// TIA Portal project "Projet Festo V4" (V20)

(* hardware
DEVICE "Station ET 200SP_1"  ET 200SP-Station
   slot 0: "Châssis_0"  Rack  6ES5 710-8MAx1
   slot 1: "6ES7512-1SK01-0AB0"  CPU 1512SP F-1 PN  6ES7 512-1SK01-0AB0  V2.8
      slot 32768: "Interface PROFINET_1"  X1
         slot 32771: "Port_3"  X1 P3
   slot 2: "F-DI 8x24VDC HF_1"  F-DI 8x24VDC HF  6ES7 136-6BA00-0CA0  V1.0
      slot 1: "F-DI 8x24VDC HF_1"  F-DI 8x24VDC HF
   slot 3: "F-DQ 4x24VDC/2A PM HF_1"  F-DQ 4x24VDC/2A PM HF  6ES7 136-6DB00-0CA0  V2.0
      slot 1: "F-DQ 4x24VDC/2A PM HF_1"  F-DQ 4x24VDC/2A PM HF
   slot 4: "F-RQ 1x24..48VDC/24..230VAC/5A_1"  F-RQ 1x24..48V DC/24..230VAC/5A  6ES7 136-6RA00-0BF0  V1.0
      slot 1: "F-RQ 1x24..48VDC/24..230VAC/5A_1"  F-RQ 1x24..48V DC/24..230VAC/5A
   slot 5: "DI 8x24VDC HF_1"  DI 8x24VDC HF  6ES7 131-6BF00-0CA0  V2.0
      slot 1: "DI 8x24VDC HF_1"  DI 8x24VDC HF
   slot 6: "DI 8x24VDC HF_2"  DI 8x24VDC HF  6ES7 131-6BF00-0CA0  V2.0
      slot 1: "DI 8x24VDC HF_2"  DI 8x24VDC HF
   slot 7: "DQ 8x24VDC/0.5A HF_1"  DQ 8x24VDC/0.5A HF  6ES7 132-6BF00-0CA0  V2.0
      slot 1: "DQ 8x24VDC/0.5A HF_1"  DQ 8x24VDC/0.5A HF
   slot 8: "DQ 8x24VDC/0.5A HF_2"  DQ 8x24VDC/0.5A HF  6ES7 132-6BF00-0CA0  V2.0
      slot 1: "DQ 8x24VDC/0.5A HF_2"  DQ 8x24VDC/0.5A HF
   slot 9: "AI 4xU/I 2-wire ST_1"  AI 4xU/I 2-wire ST  6ES7 134-6HD01-0BA1  V2.0
      slot 1: "AI 4xU/I 2-wire ST_1"  AI 4xU/I 2-wire ST
   slot 10: "AQ 4xU/I ST_1"  AQ 4xU/I ST  6ES7 135-6HD00-0BA1  V1.1
      slot 1: "AQ 4xU/I ST_1"  AQ 4xU/I ST
   slot 11: "Module serveur_1"  Server module  6ES7 193-6PA00-0AA0  V1.1
      slot 1: "Module serveur_1"  Server module
   slot 127: "BA 2xRJ45"  BA 2xRJ45  6ES7 193-6AR00-0AA0  V0.0
      slot 32769: "Port_1"  X1 P1  6ES7 193-6AR00-0AA0
      slot 32770: "Port_2"  X1 P2  6ES7 193-6AR00-0AA0
DEVICE "HMI_1"  MTP1000 Unified Comfort
   slot 0: "HMI_1"  MTP1000 Unified Comfort  6AV2 128-3KB06-0AXx  20.0.0.2
   slot 1: "HMI_RT_1"  MTP1000 Unified Comfort  6AV2 128-3KB06-0AXx  20.0.0.2
   slot 5: "HMI_1.IE_CP_1"  PROFINET Interface  20.0.0.2
      slot 1: "Interface PROFINET_1"  PROFINET Interface
         slot 1: "Port_1"  Port
         slot 2: "Port_2"  Port
   slot 6: "HMI_1.IE_CP_2"  PROFINET Interface  20.0.0.2
      slot 1: "Interface PROFINET_GBit"  PROFINET Interface
         slot 1: "Port_1"  Port
*)

// ===== PLC "6ES7512-1SK01-0AB0"  CPU 1512SP F-1 PN =====

VAR_GLOBAL   // PLC tag table "Table de variables standard"
   "Clock_Byte" AT %MB0 : Byte;   // Octet cadence B0
   "Clock_10Hz" AT %M0.0 : Bool;   // Octet cadence B0
   "Clock_5Hz" AT %M0.1 : Bool;   // Octet cadence B0
   "Clock_2.5Hz" AT %M0.2 : Bool;   // Octet cadence B0
   "Clock_2Hz" AT %M0.3 : Bool;   // Octet cadence B0
   "Clock_1.25Hz" AT %M0.4 : Bool;   // Octet cadence B0
   "Clock_1Hz" AT %M0.5 : Bool;   // Octet cadence B0
   "Clock_0.625Hz" AT %M0.6 : Bool;   // Octet cadence B0
   "Clock_0.5Hz" AT %M0.7 : Bool;   // Octet cadence B0
   "AURG_voie1" AT %I0.0 : Bool;   // Entrée Safety AURG
   "AURG_voie2" AT %I0.4 : Bool;   // Entrée Safety AURG
   "bouton_bleu" AT %I0.1 : Bool;   // acquittement apres AURG
   "voyant_bleu" AT %Q6.0 : Bool;   // Sortie Safety
   "FQ1" AT %Q6.1 : Bool;   // Sortie Safety pour relais
   "FQ2" AT %Q6.2 : Bool;   // Sortie Safety
   "libre1" AT %Q4.6 : Bool;   // free
   "libre2" AT %Q4.7 : Bool;   // free
   "libre4" AT %Q5.1 : Bool;   // free
   "libre5" AT %Q5.2 : Bool;   // free
   "libre6" AT %Q5.3 : Bool;   // free
   "libre7" AT %Q5.4 : Bool;   // free
   "libre8" AT %Q5.5 : Bool;   // free
   "Q_P_VOYANT_ROUGE" AT %Q5.6 : Bool;   // voyant rouge boite à boutons
   "Q_P_VOYANT_VERT" AT %Q5.7 : Bool;   // voyant vert boite à boutons
   "System_Byte" AT %MB1 : Byte;
   "FirstScan" AT %M1.0 : Bool;
   "DiagStatusUpdate" AT %M1.1 : Bool;
   "AlwaysTRUE" AT %M1.2 : Bool;
   "AlwaysFALSE" AT %M1.3 : Bool;
   "T_debut_bras" AT %M2.0 : Bool;
   "T_fin_bras_poste_1" AT %M2.1 : Bool;
   "T_debut_asc" AT %M2.2 : Bool;
   "T_fin_ascenseur" AT %M2.3 : Bool;
   "T_debut_test_epaisseur" AT %M2.4 : Bool;
   "Simu_VUP" AT %M20.0 : Bool;
   "Q_VUP_BR_ASC" AT %M20.1 : Bool;
   "Q_VUP_BR_MAG" AT %M20.2 : Bool;
   "I_VUP_Bras_Asc" AT %M25.1 : Bool;
   "I_VUP_Bras_Mag" AT %M25.2 : Bool;
   "I_VUP_Piece_MAG" AT %M25.3 : Bool;
   "I_VUP_Vide_Bon" AT %M25.4 : Bool;
   "Q_VUP_FAIRE_VIDE" AT %M20.3 : Bool;
   "I_VUP_Asc_Bas" AT %M25.5 : Bool;
   "I_VUP_Asc_Haut" AT %M25.6 : Bool;
   "I_VUP_Piece_Asc" AT %M25.7 : Bool;
   "Q_VUP_MONT_ASC" AT %M20.4 : Bool;
   "Q_VUP_DESC_ASC" AT %M20.5 : Bool;
   "T_debut_test_couleur" AT %M2.5 : Bool;
   "T_fin_test_couleur" AT %M2.6 : Bool;
   "T_qualite_piece" AT %MB3 : Byte;
   "T_demande_init" AT %M2.7 : Bool;   // demande d'init via IHM
   "T_fonctionnement_auto" AT %M4.6 : Bool;
   "T_fonctionnement_init" AT %M4.7 : Bool;
   "Var_Test" AT %M5.0 : Bool;
   "IHM_BRAS_MAG" AT %M5.2 : Bool;
   "IHM_BRAS_ASC" AT %M5.1 : Bool;
   "IHM_ASC_MONT" AT %M5.3 : Bool;
   "IHM_ASC_DESC" AT %M5.4 : Bool;
   "Mode_Manu_Auto" AT %M5.5 : Bool;
   "Accord_BRAS_MAG" AT %M6.1 : Bool;
   "Accord_BRAS_ASC" AT %M6.2 : Bool;
   "Accord_ASC_MONT" AT %M6.3 : Bool;
   "Accord_ASC_DESC" AT %M6.4 : Bool;
   "IHM_FAIRE_VIDE" AT %M6.5 : Bool;
   "Accord_FAIRE_VIDE" AT %M6.6 : Bool;
   "Accord_EJECTER" AT %M6.7 : Bool;
   "IHM_EJECTER" AT %M7.0 : Bool;
   "Compteurs_grande_pièce" AT %MW8 : Int;
   "Compteurs_moyenne_pièce" AT %MW10 : Int;
   "Compteurs_petite_pièce" AT %MW14 : Int;
   "IHM_Remise_a_zero" AT %M7.1 : Bool;
   "Compteurs_pièce_noire" AT %MW16 : Int;
   "Compteurs_pièce_rouge" AT %MW18 : Int;
   "Compteurs_pièce_métal" AT %MW22 : Int;
   "IHM_DEMANDE_INIT" AT %M7.2 : Bool;
   "Défaut_aspiration" AT %M7.3 : Bool;
   "Défaut_capteur_asc" AT %M7.4 : Bool;
   "Défaut_capteur_bras" AT %M7.5 : Bool;
   "IHM_ACQ_ALARMES" AT %M7.6 : Bool;
   "Compteurs_pièce_total" AT %MW26 : Int;
   "IHM_bras_animation" AT %M7.7 : Bool;
   "IHM_asc_animation" AT %M20.6 : Bool;
   "IHM_RESET_INIT" AT %M20.7 : Bool;
   "Marche_systeme" AT %M21.0 : Bool;
   "Q_VUP_EJECTER" AT %M21.1 : Bool;
   "I_VUP_Piece_Moy" AT %M21.2 : Bool;
   "I_VUP_Piece_Epais" AT %M21.3 : Bool;
   "I_VUP_Arret" AT %M21.4 : Bool;
   "I_VUP_Marche" AT %M21.5 : Bool;
   "T_Mode_Manu_VUP" AT %M21.6 : Bool;
   "I_Mode_Manu_VUP" AT %M21.7 : Bool;
END_VAR

VAR_GLOBAL   // PLC tag table "Variables T"
   "T_P_VOYANT_ROUGE" AT %M5.6 : Bool;   // voyant rouge boite à boutons
   "T_P_VOYANT_VERT" AT %M5.7 : Bool;   // voyant vert boite à boutons
   "T_Bras_Asc" AT %M12.0 : Bool;   // bras coté ascenseur
   "T_Bras_Mag" AT %M12.1 : Bool;   // bras coté magasin
   "T_Piece_Mag" AT %M12.2 : Bool;   // presence pièce magasin
   "T_Vide_Bon" AT %M12.3 : Bool;   // vide ok
   "T_Piece_Rouge" AT %M12.4 : Bool;   // capteur piece rouge/orange
   "T_Piece_Asc" AT %M12.5 : Bool;   // presence piece dans ascenceur
   "T_Piece_Metal" AT %M12.6 : Bool;   // capteur piece aluminium
   "T_Ejec_Entre" AT %M12.7 : Bool;   // verrin ejection rentré
   "T_Ejec_Sorti" AT %M13.0 : Bool;   // verrin ejection sorti
   "T_Asc_Bas" AT %M13.1 : Bool;   // ascenseur en bas
   "T_Asc_Haut" AT %M13.2 : Bool;   // ascenseur en haut
   "T_Piece_Moy" AT %M13.3 : Bool;   // capteur piece moyenne
   "T_Piece_Epais" AT %M13.4 : Bool;   // capteur piece épaisse
   "T_P_Arret" AT %M13.5 : Bool;   // bouton rouge
   "T_P_Commutateur" AT %M13.6 : Bool;   // ancien bouton aurg Festo
   "T_P_Marche" AT %M13.7 : Bool;   // bouton vert
   "T_FAIRE_VIDE" AT %M4.0 : Bool;   // monostable faire vide
   "T_BR_ASC" AT %M4.1 : Bool;   // bistable bras vers ascenseur
   "T_BR_MAG" AT %M4.2 : Bool;   // bistable bras vers mag
   "T_EJECTER" AT %M4.3 : Bool;   // monostable ejection piece
   "T_MONT_ASC" AT %M4.4 : Bool;   // bistable monter ascenseur
   "T_DESC_ASC" AT %M4.5 : Bool;   // bistable descendre ascenseur
   "T_Fin_test_epaisseur" AT %M6.0 : Bool;
END_VAR

VAR_GLOBAL   // PLC tag table "Var I/Q"
   "I_Bras_Asc" AT %I12.0 : Bool;   // bras coté ascenseur
   "I_Bras_Mag" AT %I12.1 : Bool;   // bras coté magasin
   "I_Piece_Mag" AT %I12.2 : Bool;   // presence pièce magasin
   "I_Vide_Bon" AT %I12.3 : Bool;   // vide ok
   "I_Piece_Rouge" AT %I12.4 : Bool;   // capteur piece rouge/orange
   "I_Piece_Asc" AT %I12.5 : Bool;   // presence piece dans ascenceur
   "I_Piece_Metal" AT %I12.6 : Bool;   // capteur piece aluminium
   "I_Ejec_Entre" AT %I12.7 : Bool;   // verrin ejection rentré
   "I_Ejec_Sorti" AT %I13.0 : Bool;   // verrin ejection sorti
   "I_Asc_Bas" AT %I13.1 : Bool;   // ascenseur en bas
   "I_Asc_Haut" AT %I13.2 : Bool;   // ascenseur en haut
   "I_Piece_Moy" AT %I13.3 : Bool;   // capteur piece moyenne
   "I_Piece_Epais" AT %I13.4 : Bool;   // capteur piece épaisse
   "I_P_Arret" AT %I13.5 : Bool;   // bouton rouge
   "I_P_Commutateur" AT %I13.6 : Bool;   // ancien bouton aurg Festo
   "I_P_Marche" AT %I13.7 : Bool;   // bouton vert
   "Q_FAIRE_VIDE" AT %Q5.0 : Bool;   // monostable faire vide
   "Q_BR_ASC" AT %Q4.0 : Bool;   // bistable bras vers ascenseur
   "Q_BR_MAG" AT %Q4.1 : Bool;   // bistable bras vers mag
   "Q_EJECTER" AT %Q4.2 : Bool;   // monostable ejection piece
   "Q_MONT_ASC" AT %Q4.3 : Bool;   // bistable monter ascenseur
   "Q_DESC_ASC" AT %Q4.4 : Bool;   // bistable descendre ascenseur
END_VAR

// folder: DB

DATA_BLOCK "Marche_Arret_DB"   // DB3
{ S7_Optimized_Access := 'TRUE' }
VERSION : 0.1
// stored: InstanceOfName Marche_Arret
"Marche_Arret"
BEGIN
END_DATA_BLOCK

DATA_BLOCK "Bras_poste_1_DB"   // DB4
{ S7_Optimized_Access := 'TRUE' }
VERSION : 0.1
// stored: InstanceOfName Bras_poste_1
"Bras_poste_1"
BEGIN
END_DATA_BLOCK

DATA_BLOCK "Ascenseur_poste_1_DB"   // DB5
{ S7_Optimized_Access := 'TRUE' }
VERSION : 0.1
// stored: InstanceOfName Ascenseur_poste_1
"Ascenseur_poste_1"
BEGIN
END_DATA_BLOCK

DATA_BLOCK "Test_Épaisseur_DB"   // DB6
{ S7_Optimized_Access := 'TRUE' }
VERSION : 0.1
// stored: InstanceOfName Test_Épaisseur
"Test_Épaisseur"
BEGIN
END_DATA_BLOCK

DATA_BLOCK "Conduite_DB"   // DB7
{ S7_Optimized_Access := 'TRUE' }
VERSION : 0.1
// stored: InstanceOfName Conduite
"Conduite"
BEGIN
END_DATA_BLOCK

DATA_BLOCK "Test_couleur_DB"   // DB8
{ S7_Optimized_Access := 'TRUE' }
VERSION : 0.1
// stored: InstanceOfName Test_couleur
"Test_couleur"
BEGIN
END_DATA_BLOCK

DATA_BLOCK "Initialisation_DB"   // DB9
{ S7_Optimized_Access := 'TRUE' }
VERSION : 0.1
// stored: InstanceOfName Initialisation
"Initialisation"
BEGIN
END_DATA_BLOCK

DATA_BLOCK "Mode_Manu_DB"   // DB10
{ S7_Optimized_Access := 'TRUE' }
VERSION : 0.1
// stored: InstanceOfName Mode_Manu
"Mode_Manu"
BEGIN
END_DATA_BLOCK

DATA_BLOCK "Compteurs_DB"   // DB11
{ S7_Optimized_Access := 'TRUE' }
VERSION : 0.1
// stored: InstanceOfName Compteurs
"Compteurs"
BEGIN
END_DATA_BLOCK

DATA_BLOCK "Alarmes_DB"   // DB12
{ S7_Optimized_Access := 'TRUE' }
VERSION : 0.1
// stored: InstanceOfName Alarmes
"Alarmes"
BEGIN
END_DATA_BLOCK

DATA_BLOCK "Default_SupervisionDB"   // DB13
{ S7_Optimized_Access := 'TRUE' }
VERSION : 0.1
// stored: InstanceOfName Default_SupervisionFB
"Default_SupervisionFB"
BEGIN
END_DATA_BLOCK

DATA_BLOCK "IHM_DB"   // DB14
{ S7_Optimized_Access := 'TRUE' }
VERSION : 0.1
// stored: InstanceOfName IHM
"IHM"
BEGIN
END_DATA_BLOCK

// folder: Safety

DATA_BLOCK "Main_Safety_RTG1_DB"   // DB1, F_DB
{ S7_Optimized_Access := 'TRUE' }
NAME : FUSI
VERSION : 0.1
// stored: InstanceOfName Main_Safety_RTG1
"Main_Safety_RTG1"
BEGIN
END_DATA_BLOCK

DATA_BLOCK "Arret_Urgence_DB"   // DB2, F_DB
{ S7_Optimized_Access := 'TRUE' }
VERSION : 0.1
// stored: InstanceOfName Arret_Urgence
"Arret_Urgence"
BEGIN
END_DATA_BLOCK

// folder: (top level)

FUNCTION_BLOCK "Test_Épaisseur"   // FB3, SCL
{ S7_Optimized_Access := 'TRUE' }
VERSION : 0.1
   VAR_INPUT
      asc_haut : Bool;
      capteur_moy : Bool;
      capteur_grd : Bool;
      asc_bas : Bool;
      presence_piece_asc : Bool;
      marche : Bool;
   END_VAR
   VAR_OUTPUT
      DESC_ASC : Bool;
      EJECTER : Bool;
      FIN_TEST : Bool;
   END_VAR
   VAR
      Etape_Test_epaisseur : Int;
      CE100_110 : Bool;
      CE110_120 : Bool;
      CE130_100 : Bool;
      CE140_100 : Bool;
      CE150_100 : Bool;
      CE120_130 : Bool;
      CE120_140 : Bool;
      CE120_150 : Bool;
      Timer_test_pièce : TON_TIME;
      CE140_145 : Bool;
      CE150_155 : Bool;
      CE130_140 : Bool;
      CE150_160 : Bool;
      CE170_180 : Bool;
      "#CE140_100" : Bool;
      CE160_100 : Bool;
      CE180_100 : Bool;
      CE120_170 : Bool;
      CE140_190 : Bool;
      CE160_190 : Bool;
      CE180_190 : Bool;
      CE190_100 : Bool;
      Timer_ejecte_pièce : TON_TIME;
      Timer_fin_test : TON_TIME;
   END_VAR
BEGIN
   #Timer_test_pièce(IN:=#Etape_Test_epaisseur=110,PT:=T#1s);
   #Timer_ejecte_pièce(IN := #Etape_Test_epaisseur = 140 OR #Etape_Test_epaisseur = 150 OR #Etape_Test_epaisseur = 180,
                       PT := T#500ms);
   #Timer_fin_test(IN := #Etape_Test_epaisseur = 190,
                     PT := T#1s);

   #CE100_110 := #Etape_Test_epaisseur = 100 AND #asc_haut AND #marche;
   #CE110_120 := #Etape_Test_epaisseur = 110 AND #Timer_test_pièce.Q;
   //Grande Pièce
   #CE120_130 := #Etape_Test_epaisseur = 120 AND #capteur_moy AND #capteur_grd;
   #CE130_140 := #Etape_Test_epaisseur = 130 AND #asc_bas;
   #CE140_190 := #Etape_Test_epaisseur = 140 AND NOT #presence_piece_asc AND #Timer_ejecte_pièce.Q;
   //Moyenne Pièce
   #CE120_150 := #Etape_Test_epaisseur = 120 AND #capteur_moy AND NOT #capteur_grd;
   #CE150_160 := #Etape_Test_epaisseur = 150 AND NOT #presence_piece_asc AND #Timer_ejecte_pièce.Q;
   #CE160_190 := #Etape_Test_epaisseur = 160 AND #asc_bas;
   //Petite Pièce
   #CE120_170 := #Etape_Test_epaisseur = 120 AND NOT #capteur_moy AND NOT #capteur_grd;
   #CE170_180 := #Etape_Test_epaisseur = 170 AND #asc_bas;
   #CE180_190 := #Etape_Test_epaisseur = 180 AND NOT #presence_piece_asc AND #Timer_ejecte_pièce.Q;
   //Fin TEST
   #CE190_100 := #Etape_Test_epaisseur = 190 AND #Timer_fin_test.Q;

   IF #CE100_110 THEN
       #Etape_Test_epaisseur := 110;
   END_IF;

   IF #CE110_120 THEN
       #Etape_Test_epaisseur := 120;
   END_IF;

   IF #CE120_130 THEN
       #Etape_Test_epaisseur := 130;
   END_IF;

   IF #CE130_140 THEN
       #Etape_Test_epaisseur := 140;
   END_IF;

   IF #CE140_190 THEN
       #Etape_Test_epaisseur := 190;
   END_IF;

   IF #CE120_150 THEN
       #Etape_Test_epaisseur := 150;
   END_IF;

   IF #CE150_160 THEN
       #Etape_Test_epaisseur := 160;
   END_IF;

   IF #CE160_190 THEN
       #Etape_Test_epaisseur := 190;
   END_IF;

   IF #CE120_170 THEN
       #Etape_Test_epaisseur := 170;
   END_IF;

   IF #CE170_180 THEN
       #Etape_Test_epaisseur := 180;
   END_IF;

   IF #CE180_190 THEN
       #Etape_Test_epaisseur := 190;
   END_IF;

   IF #CE190_100 THEN
       #Etape_Test_epaisseur := 100;
   END_IF;




   #FIN_TEST := #Etape_Test_epaisseur = 190;
END_FUNCTION_BLOCK

FUNCTION_BLOCK "Marche_Arret"   // FB4, SCL
{ S7_Optimized_Access := 'TRUE' }
VERSION : 0.1
   VAR_INPUT
      Bouton_Rouge : Bool;
      Bouton_Vert : Bool;
   END_VAR
   VAR_OUTPUT
      Voyant_vert : Bool;
      Marche_systeme : Bool;
      Voyant_rouge : Bool;
   END_VAR
   VAR
      Etape_Marche_Arret : Int;
      CE10_20 : Bool;
      CE20_10 : Bool;
   END_VAR
BEGIN
   //Fonctionnement du marche arret
   //Lance un cycle si le bouton vert est appuyer et arrete si le rouge est appuyer


   #CE10_20 := #Etape_Marche_Arret = 10 AND #Bouton_Vert AND NOT #Bouton_Rouge;
   #CE20_10 := #Etape_Marche_Arret = 20 AND #Bouton_Rouge;

   IF #CE10_20 THEN
       #Etape_Marche_Arret := 20;
   END_IF;
   IF #CE20_10 THEN
       #Etape_Marche_Arret := 10;
   END_IF;

   #Voyant_vert := #Etape_Marche_Arret = 20;
   #Voyant_rouge := #Etape_Marche_Arret = 10;
   #Marche_systeme := #Etape_Marche_Arret = 20;
END_FUNCTION_BLOCK

FUNCTION_BLOCK "Bras_poste_1"   // FB5, SCL
{ S7_Optimized_Access := 'TRUE' }
VERSION : 0.1
   VAR_INPUT
      bras_asc : Bool;
      presence_piece : Bool;
      marche : Bool;
      bras_mag : Bool;
      vide_bon : Bool;
   END_VAR
   VAR_OUTPUT
      FIN_BRAS_POSTE_1 : Bool;
   END_VAR
   VAR
      Etape_Bras_Poste_1 : Int;
      CE400_410 : Bool;
      CE410_420 : Bool;
      CE420_430 : Bool;
      CE430_440 : Bool;
      CE440_450 : Bool;
      CE450_400 : Bool;
      CE450_410 : Bool;
      Timer_fin_bras : TON_TIME;
      CE450_460 : Bool;
      CE460_410 : Bool;
      CE460_400 : Bool;
   END_VAR
BEGIN
   //Fonctionnement du cycle du bras

   //Timer de fin de cycle bras pas sécurité
   #Timer_fin_bras(IN:=#Etape_Bras_Poste_1=460,PT:=T#1s);

   //Conditions d'évolutions
   #CE400_410 := #Etape_Bras_Poste_1 = 400 AND #presence_piece AND #marche;
   #CE410_420 := #Etape_Bras_Poste_1 = 410 AND #bras_mag;
   #CE420_430 := #Etape_Bras_Poste_1 = 420 AND #vide_bon;
   #CE430_440 := #Etape_Bras_Poste_1 = 430 AND #bras_asc;
   #CE440_450 := #Etape_Bras_Poste_1 = 440 AND NOT #vide_bon;
   #CE450_460 := #Etape_Bras_Poste_1 = 450 AND #bras_mag;
   #CE460_400 := #Etape_Bras_Poste_1 = 460 AND #Timer_fin_bras.Q;

   IF #CE400_410 THEN
       #Etape_Bras_Poste_1 := 410;
   END_IF;

   IF #CE410_420 THEN
       #Etape_Bras_Poste_1 := 420;
   END_IF;

   IF #CE420_430 THEN
       #Etape_Bras_Poste_1 := 430;
   END_IF;

   IF #CE430_440 THEN
       #Etape_Bras_Poste_1 := 440;
   END_IF;

   IF #CE440_450 THEN
       #Etape_Bras_Poste_1 := 450;
   END_IF;

   IF #CE450_460 THEN
       #Etape_Bras_Poste_1 := 460;
   END_IF;

   IF #CE460_400 THEN
       #Etape_Bras_Poste_1 := 400;
   END_IF;

   //Fin cycle bras pour G7 de conduite
   #FIN_BRAS_POSTE_1 := #Etape_Bras_Poste_1 = 460;
END_FUNCTION_BLOCK

FUNCTION_BLOCK "Test_couleur"   // FB6, SCL
{ S7_Optimized_Access := 'TRUE' }
VERSION : 0.1
   VAR_INPUT
      marche : Bool;
      piece_rouge : Bool;
      piece_metal : Bool;
      Ejecteur_sortie : Bool;
   END_VAR
   VAR_OUTPUT
      Qualite_piece : Byte;
      Fin_test_couleur : Bool;
   END_VAR
   VAR
      Timer_test_couleur : TON_TIME;
      Timer_fin_test_couleur : TON_TIME;
      Etape_test_couleur : Int;
      CE700_710 : Bool;
      CE710_720 : Bool;
      CE720_700 : Bool;
      CE720_730 : Bool;
      CE730_740 : Bool;
      CE730_750 : Bool;
      CE730_760 : Bool;
      CE740_700 : Bool;
      CE750_700 : Bool;
      CE760_700 : Bool;
   END_VAR
BEGIN
   #Timer_test_couleur(IN:=#Etape_test_couleur=710,
                       PT:=T#1s);
   #Timer_fin_test_couleur(IN:=#Etape_test_couleur=720,
                           PT:=T#1s);

   #CE700_710 := #Etape_test_couleur = 700 AND #marche;
   #CE710_720 := #Etape_test_couleur = 710 AND #Timer_test_couleur.Q;
   #CE720_730 := #Etape_test_couleur = 720 AND #Timer_fin_test_couleur.Q;

   #CE730_740 := #Etape_test_couleur = 730 AND #piece_rouge AND NOT #piece_metal ; //piece rouge
   #CE730_750 := #Etape_test_couleur = 730 AND #piece_metal; //piece métal
   #CE730_760 := #Etape_test_couleur = 730 AND NOT #piece_metal AND NOT #piece_rouge; //piece noire

   #CE740_700 := #Etape_test_couleur = 740 AND #Ejecteur_sortie;
   #CE750_700 := #Etape_test_couleur = 750 AND #Ejecteur_sortie;
   #CE760_700 := #Etape_test_couleur = 760 AND #Ejecteur_sortie;

   IF #CE700_710 THEN
       #Etape_test_couleur := 710;
   END_IF;
   IF #CE710_720 THEN
       #Etape_test_couleur := 720;
   END_IF;
   IF #CE720_730 THEN
       #Etape_test_couleur := 730;
   END_IF;
   IF #CE730_740 THEN
       #Etape_test_couleur := 740;
   END_IF;
   IF #CE730_750 THEN
       #Etape_test_couleur := 750;
   END_IF;
   IF #CE730_760 THEN
       #Etape_test_couleur := 760;
   END_IF;
   IF #CE740_700 THEN
       #Etape_test_couleur := 700;
   END_IF;
   IF #CE750_700 THEN
       #Etape_test_couleur := 700;
   END_IF;
   IF #CE760_700 THEN
       #Etape_test_couleur := 700;
   END_IF;




   #Fin_test_couleur := #Etape_test_couleur = 720;
END_FUNCTION_BLOCK

FUNCTION_BLOCK "Ascenseur_poste_1"   // FB7, SCL
{ S7_Optimized_Access := 'TRUE' }
VERSION : 0.1
   VAR_INPUT
      asc_bas : Bool;
      presence_piece_asc : Bool;
      asc_haut : Bool;
      Fin_test_epaisseur : Bool;
      marche : Bool;
   END_VAR
   VAR_OUTPUT
      MONTER_ASC : Bool;
      DESCENDRE_ASC : Bool;
      FIN_ASCENSEUR : Bool;
   END_VAR
   VAR
      Etape_Ascenseur : Int;
      CE500_510 : Bool;
      CE510_520 : Bool;
      CE520_530 : Bool;
      CE530_500 : Bool;
      Timer_fin_asc : TON_TIME;
      CE530_540 : Bool;
      CE540_500 : Bool;
   END_VAR
BEGIN
   //Fonctionnement de l'ascenseur

   //Timer de fin de cycle de l'ascenseur par sécurité
   #Timer_fin_asc(IN:=#Etape_Ascenseur=540,
                  PT:=T#1s);

   //Conditions d'évolutions
   #CE500_510 := #Etape_Ascenseur = 500 AND #asc_bas AND #presence_piece_asc AND #marche; //Lancement du fct ASC si le G7 de conduite le permet
   #CE510_520 := #Etape_Ascenseur = 510 AND #asc_haut;
   #CE520_530 := #Etape_Ascenseur = 520 AND #Fin_test_epaisseur;
   #CE530_540 := #Etape_Ascenseur = 530 AND #asc_bas;
   #CE540_500 := #Etape_Ascenseur = 540 AND #Timer_fin_asc.Q;

   IF #CE500_510 THEN
       #Etape_Ascenseur := 510;
   END_IF;

   IF #CE510_520 THEN
       #Etape_Ascenseur := 520;
   END_IF;

   IF #CE520_530 THEN
       #Etape_Ascenseur := 530;
   END_IF;

   IF #CE530_540 THEN
       #Etape_Ascenseur := 540;
   END_IF;

   IF #CE540_500 THEN
       #Etape_Ascenseur := 500;
   END_IF;

   //Fin cycle ascenseur pour G7 de conduite
   #FIN_ASCENSEUR := #Etape_Ascenseur = 540;
END_FUNCTION_BLOCK

FUNCTION_BLOCK "Conduite"   // FB8, SCL
{ S7_Optimized_Access := 'TRUE' }
VERSION : 0.1
   VAR_INPUT
      Marche : Bool;
      Fin_bras : Bool;
      Fin_ascenseur : Bool;
      Fin_test_couleur : Bool;
      Fin_test_epaisseur : Bool;
      Fonctionnement_init : Bool;
      présence_pice_mag : Bool;
   END_VAR
   VAR_OUTPUT
      DEBUT_BRAS : Bool;
      DEBUT_ASCENSEUR : Bool;
      DEBUT_EPAISSEUR : Bool;
      DEBUT_TEST_COULEUR : Bool;
      fonctionnement_auto : Bool;
   END_VAR
   VAR
      CE1000_1010 : Bool;
      CE1010_1020 : Bool;
      CE1020_1030 : Bool;
      CE1030_1000 : Bool;
      CE1030_1010 : Bool;
      Etape_conduite : Int;
      CE1020_1025 : Bool;
      CE1025_1030 : Bool;
   END_VAR
BEGIN
   //G7 de conduite, lance les autres G7

   #CE1000_1010 := #Etape_conduite = 1000 AND #Marche AND NOT #Fonctionnement_init AND #présence_pice_mag;
   #CE1010_1020 := #Etape_conduite = 1010 AND #Fin_bras;
   #CE1020_1025 := #Etape_conduite = 1020 AND #Fin_test_couleur;
   #CE1025_1030 := #Etape_conduite = 1025 AND #Fin_test_epaisseur;
   #CE1030_1000 := #Etape_conduite = 1030 AND #Fin_ascenseur;

   IF #CE1000_1010 THEN
       #Etape_conduite := 1010;
   END_IF;

   IF #CE1010_1020 THEN
       #Etape_conduite := 1020;
   END_IF;

   IF #CE1020_1025 THEN
       #Etape_conduite := 1025;
   END_IF;

   IF #CE1025_1030 THEN
       #Etape_conduite := 1030;
   END_IF;

   IF #CE1030_1000 THEN
       #Etape_conduite := 1000;
   END_IF;

   #DEBUT_BRAS := #Etape_conduite = 1010;
   #DEBUT_TEST_COULEUR := #Etape_conduite = 1020;
   #DEBUT_ASCENSEUR := #Etape_conduite = 1025;
   #DEBUT_EPAISSEUR := #Etape_conduite = 1025;

   #fonctionnement_auto := #Etape_conduite = 1010 OR #Etape_conduite = 1020 OR #Etape_conduite = 1030 OR #Etape_conduite=1025;

   IF "T_fonctionnement_auto" THEN
       "Accord_ASC_DESC" := FALSe;
       "Accord_ASC_MONT" := FALSe;
       "Accord_BRAS_ASC" := FALSe;
       "Accord_BRAS_MAG" := FALSe;
       "Accord_EJECTER" := FALSe;
       "Accord_FAIRE_VIDE" := FALSe;
   END_IF;
END_FUNCTION_BLOCK

FUNCTION_BLOCK "Initialisation"   // FB9, SCL
{ S7_Optimized_Access := 'TRUE' }
VERSION : 0.1
   VAR_INPUT
      Bras_asc : Bool;
      Asc_bas : Bool;
      Bras_mag : Bool;
      Demande_init : Bool;
      fonctionnement_auto : Bool;
      IHM_DEMANDE_INIT : Bool;
   END_VAR
   VAR_OUTPUT
      BR_MAG : Bool;
      DESC_ASC : Bool;
      BR_ASC : Bool;
      Fonctionnement_init : Bool;
   END_VAR
   VAR
      CE2000_2010 : Bool;
      CE2010_2020 : Bool;
      CE2020_2030 : Bool;
      CE2030_2000 : Bool;
      Etape_init : Int;
      CE2030_2040 : Bool;
      CE2040_2000 : Bool;
   END_VAR
BEGIN
   //Fonctionnement de l'initialisation
   //Lancer par une entrée IHM
   //
   #CE2000_2010 := #Etape_init = 2000 AND #IHM_DEMANDE_INIT AND NOT #fonctionnement_auto;
   #CE2010_2020 := #Etape_init = 2010 AND #Bras_mag;
   #CE2020_2030 := #Etape_init = 2020 AND #Asc_bas;
   #CE2030_2000 := #Etape_init = 2030 AND #Bras_asc;

   IF #CE2000_2010 THEN
       #Etape_init := 2010;
   END_IF;
   IF #CE2010_2020 THEN
       #Etape_init := 2020;
   END_IF;
   IF #CE2020_2030 THEN
       #Etape_init := 2030;
   END_IF;
   IF #CE2030_2000 THEN
       #Etape_init := 2000;
   END_IF;






   //Informe que le système effectue une init 
   #Fonctionnement_init := #Etape_init = 2010 OR #Etape_init = 2020 OR #Etape_init = 2030;
END_FUNCTION_BLOCK

FUNCTION_BLOCK "Mode_Manu"   // FB10, SCL
{ S7_Optimized_Access := 'TRUE' }
VERSION : 0.1
   VAR_INPUT
      IHM_EJECTER : Bool;
      IHM_Bras_MAG : Bool;
      IHM_BRAS_ASC : Bool;
      IHM_ASC_MONT : Bool;
      IHM_ASc_DESC : Bool;
      IHM_FAIRE_VIDE : Bool;
   END_VAR
   VAR_OUTPUT
      Accord_EJECTER : Bool;
      Accord_BRAS_MAG : Bool;
      Accord_ASC_MONT : Bool;
      Accord_ASC_BAS : Bool;
      Accord_FAIRE_VIDE : Bool;
   END_VAR
   VAR_IN_OUT
      Accord_BRAS_ASC : Bool;
   END_VAR
BEGIN
   IF #IHM_Bras_MAG AND NOT "T_Asc_Haut"  AND NOT #IHM_BRAS_ASC THEN
       #Accord_BRAS_MAG := TRUE;
       #Accord_BRAS_ASC := FALSE;
   END_IF;

   IF #IHM_BRAS_ASC AND NOT "T_Asc_Haut" AND NOT #IHM_Bras_MAG THEN
       #Accord_BRAS_ASC := TRUE;
       #Accord_BRAS_MAG := FALSE;
   END_IF;

   IF #IHM_ASC_MONT AND NOT "T_Bras_Asc" AND NOT #Accord_BRAS_ASC THEN
       #Accord_ASC_MONT := TRUE;
       #Accord_ASC_BAS := FALSE;
   END_IF;

   IF #IHM_ASc_DESC AND NOT "T_Bras_Asc" THEN
       #Accord_ASC_MONT := FALSE;
       #Accord_ASC_BAS := TRUE;
   END_IF;

   IF #IHM_FAIRE_VIDE THEN
       #Accord_FAIRE_VIDE := TRUE;
   END_IF;
   IF NOT #IHM_FAIRE_VIDE THEN
       #Accord_FAIRE_VIDE := FALSE;
   END_IF;

   IF #IHM_EJECTER THEN
       #Accord_EJECTER := TRUE;
   END_IF;
   IF NOT #IHM_EJECTER THEN
       #Accord_EJECTER := FALSE;
   END_IF;


   IF "IHM_RESET_INIT" THEN
       #Accord_ASC_BAS := FALSE;
       #Accord_ASC_MONT := FALSE;
       #Accord_BRAS_ASC := FALSE;
       #Accord_BRAS_MAG := FALSE;
       #Accord_EJECTER := FALSE;
       #Accord_FAIRE_VIDE := FALSE;
   END_IF;
END_FUNCTION_BLOCK

FUNCTION_BLOCK "Compteurs"   // FB11, SCL
{ S7_Optimized_Access := 'TRUE' }
VERSION : 0.1
   VAR_INPUT
      IHM_Remise_a_zero : Bool;
   END_VAR
   VAR
      R_trig_grande_p : R_TRIG;
      R_trig_petite_p : R_TRIG;
      R_trig_moyenne_p : R_TRIG;
      R_trig_noire_p : R_TRIG;
      R_trig_rouge_p : R_TRIG;
      R_trig_métal_p : R_TRIG;
   END_VAR
BEGIN
   //Taille des pièces
   #R_trig_grande_p(CLK:="Test_Épaisseur_DB".Etape_Test_epaisseur = 170);
   #R_trig_petite_p(CLK := "Test_Épaisseur_DB".Etape_Test_epaisseur = 130);
   #R_trig_moyenne_p(CLK:="Test_Épaisseur_DB".Etape_Test_epaisseur = 150);

   //Couleurs des pièces
   #R_trig_noire_p(CLK := "Test_couleur_DB".Etape_test_couleur = 760);
   #R_trig_rouge_p(CLK := "Test_couleur_DB".Etape_test_couleur = 740);
   #R_trig_métal_p(CLK := "Test_couleur_DB".Etape_test_couleur = 750);

   //Condition d'incrémentation taille
   IF #R_trig_grande_p.Q THEN
       "Compteurs_grande_pièce" := "Compteurs_grande_pièce" + 1;
   END_IF;
   IF #R_trig_moyenne_p.Q THEN
       "Compteurs_moyenne_pièce" := "Compteurs_moyenne_pièce" + 1;
   END_IF;
   IF #R_trig_petite_p.Q THEN
       "Compteurs_petite_pièce" := "Compteurs_petite_pièce" + 1;
   END_IF;
   //Condition d'incrémentation couleur
   IF #R_trig_noire_p.Q THEN
       "Compteurs_pièce_noire" := "Compteurs_pièce_noire" + 1;
   END_IF;
   IF #R_trig_rouge_p.Q THEN
       "Compteurs_pièce_rouge" := "Compteurs_pièce_noire" + 1;
   END_IF;
   IF #R_trig_métal_p.Q THEN
       "Compteurs_pièce_métal" := "Compteurs_pièce_métal" + 1;
   END_IF;

   //Pièce total
   "Compteurs_pièce_total" := "Compteurs_pièce_noire" + "Compteurs_pièce_noire" + "Compteurs_pièce_métal" + "Compteurs_grande_pièce" + "Compteurs_moyenne_pièce" + "Compteurs_petite_pièce";

   //RAZ compteurs
   IF #IHM_Remise_a_zero THEN
       "Compteurs_grande_pièce" := 0;
       "Compteurs_moyenne_pièce" := 0;
       "Compteurs_petite_pièce" := 0;
       "Compteurs_pièce_noire" := 0;
       "Compteurs_pièce_rouge" := 0;
       "Compteurs_pièce_métal" := 0;
       "Compteurs_pièce_total" := 0;
   END_IF;
END_FUNCTION_BLOCK

FUNCTION_BLOCK "Alarmes"   // FB12, SCL
{ S7_Optimized_Access := 'TRUE' }
VERSION : 0.1
   VAR_INPUT
      Faire_vide : Bool;
      vide_bon : Bool;
      Asc_haut : Bool;
      Asc_bas : Bool;
      IHM_ACQ_ALARMES : Bool;
      Bras_mag : Bool;
      Bras_asc : Bool;
   END_VAR
   VAR_OUTPUT
      Defaut_aspiration : Bool;
      Defaut_capteur_asc : Bool;
      Defaut_capteurs_bras : Bool;
   END_VAR
   VAR
      Timer_defaut_aspiration : TON_TIME;
   END_VAR
BEGIN
   //Gestion des défauts et alarmes

   //Temps avant défaut de l'aspiration
   #Timer_defaut_aspiration(IN := #Faire_vide AND NOT #vide_bon,
                            PT := T#4s);

   //Création des défauts selon certaines conditions.
   IF #Timer_defaut_aspiration.Q THEN //Défauta aspiration
       #Defaut_aspiration := TRUE;

   END_IF;
   IF #Asc_haut AND #Asc_bas THEN //Défaut des capteurs de l'ascenseur
       #Defaut_capteur_asc := TRUE;
   END_IF;
   IF #Bras_mag AND #Bras_asc THEN//Défaut des capteurs du bras
       #Defaut_capteurs_bras := TRUE;
   END_IF;


   //Acquitement des alarmes
   IF #IHM_ACQ_ALARMES THEN
       #Defaut_aspiration:= FALSE;
       #Defaut_capteur_asc := FALSE;
       #Defaut_capteurs_bras := FALSE;
   END_IF;
END_FUNCTION_BLOCK

FUNCTION_BLOCK "Default_SupervisionFB"   // FB13, ProDiag
{ S7_Optimized_Access := 'TRUE' }
   VAR
      PC_Flags : PC_Flags_V2;
      State : SV_FB_State_V2;
   END_VAR
   VAR_TEMP
      t_TempSvStateUDT : SV_State_V2;
      t_TempAlarmInstance : <type 200004f>;
      t_TempAsocValue1 : Variant;
      t_TempAsocValue2 : Variant;
      t_TempAsocValue3 : Variant;
   END_VAR
BEGIN
END_FUNCTION_BLOCK

FUNCTION "Sortie" : Void   // FC5, SCL
{ S7_Optimized_Access := 'TRUE' }
VERSION : 0.1
BEGIN
   //Rassemblement des T reliés aux sorties
   "T_FAIRE_VIDE" := "Bras_poste_1_DB".Etape_Bras_Poste_1 = 420 OR "Bras_poste_1_DB".Etape_Bras_Poste_1 = 430 OR "Mode_Manu_DB".Accord_FAIRE_VIDE;
   "T_BR_ASC" := "Bras_poste_1_DB".Etape_Bras_Poste_1 = 430 OR "Initialisation_DB".Etape_init = 2030 OR "Accord_BRAS_ASC";
   "T_BR_MAG" := "Bras_poste_1_DB".Etape_Bras_Poste_1= 410 OR "Bras_poste_1_DB".Etape_Bras_Poste_1= 450 OR "Initialisation_DB".Etape_init = 2010 OR "Accord_BRAS_MAG";
   "T_EJECTER" := "Test_Épaisseur_DB".Etape_Test_epaisseur = 140 OR "Test_Épaisseur_DB".Etape_Test_epaisseur = 150 OR "Test_Épaisseur_DB".Etape_Test_epaisseur = 180 OR "Accord_EJECTER";
   IF NOT "Simu_VUP" THEN

       "T_MONT_ASC" := "Ascenseur_poste_1_DB".Etape_Ascenseur = 510 OR "Accord_ASC_MONT";

   END_IF;
   IF "Simu_VUP" THEN

       "T_MONT_ASC" := "Ascenseur_poste_1_DB".Etape_Ascenseur = 510 OR "Ascenseur_poste_1_DB".Etape_Ascenseur = 520 OR "Accord_ASC_MONT";

   END_IF;
   "T_DESC_ASC" := "Ascenseur_poste_1_DB".Etape_Ascenseur = 530 OR "Test_Épaisseur_DB".Etape_Test_epaisseur = 130 OR "Test_Épaisseur_DB".Etape_Test_epaisseur = 160 OR "Test_Épaisseur_DB".Etape_Test_epaisseur = 170 OR "Accord_ASC_DESC" OR "Initialisation_DB".Etape_init=2020;
END_FUNCTION

ORGANIZATION_BLOCK "Main"   // OB1, LAD, ProgramCycle
TITLE = "Main Program Sweep (Cycle)"
{ S7_Optimized_Access := 'TRUE' }
VERSION : 0.1
   VAR_INPUT
      Initial_Call : Bool;   // Initial call of this OB
      Remanence : Bool;   // =True, if remanent data are available
   END_VAR
BEGIN

REGION Network 1: IDDI en mode réel
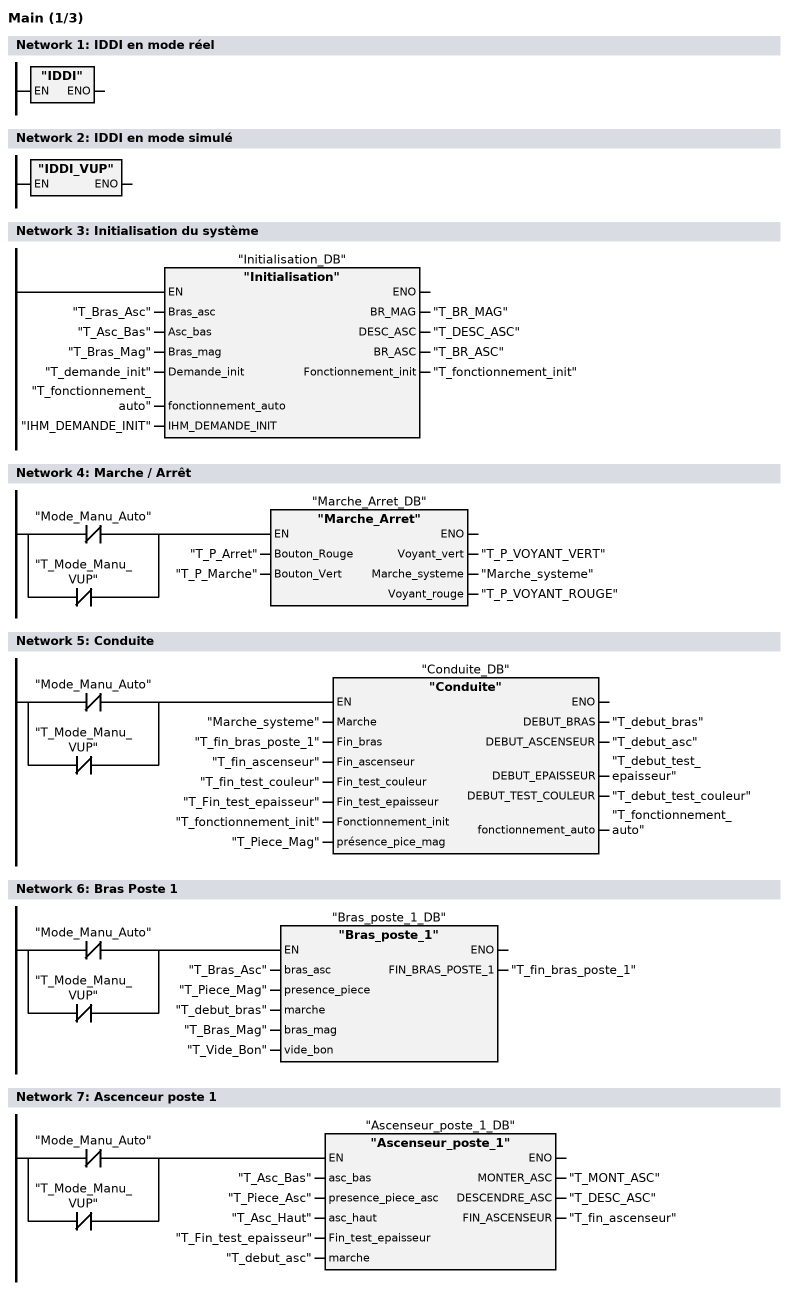
   RUNG wire#powerrail
      "IDDI"()
   END_RUNG
   // the same network as SCL:
   "IDDI"();
END_REGION

REGION Network 2: IDDI en mode simulé
   RUNG wire#powerrail
      "IDDI_VUP"()
   END_RUNG
   // the same network as SCL:
   "IDDI_VUP"();
END_REGION

REGION Network 3: Initialisation du système
   RUNG wire#powerrail
      "Initialisation_DB"(Bras_asc := "T_Bras_Asc", Asc_bas := "T_Asc_Bas", Bras_mag := "T_Bras_Mag", Demande_init := "T_demande_init", fonctionnement_auto := "T_fonctionnement_auto", IHM_DEMANDE_INIT := "IHM_DEMANDE_INIT", BR_MAG => "T_BR_MAG", DESC_ASC => "T_DESC_ASC", BR_ASC => "T_BR_ASC", Fonctionnement_init => "T_fonctionnement_init")
   END_RUNG
   // the same network as SCL:
   "Initialisation_DB"(Bras_asc := "T_Bras_Asc",   // "Initialisation"
                       Asc_bas := "T_Asc_Bas",
                       Bras_mag := "T_Bras_Mag",
                       Demande_init := "T_demande_init",
                       fonctionnement_auto := "T_fonctionnement_auto",
                       IHM_DEMANDE_INIT := "IHM_DEMANDE_INIT",
                       BR_MAG => "T_BR_MAG",
                       DESC_ASC => "T_DESC_ASC",
                       BR_ASC => "T_BR_ASC",
                       Fonctionnement_init => "T_fonctionnement_init");
END_REGION

REGION Network 4: Marche / Arrêt
   RUNG wire#powerrail
      I_Contact( "Mode_Manu_Auto" )
      wire#w1
      "Marche_Arret_DB"(Bouton_Rouge := "T_P_Arret", Bouton_Vert := "T_P_Marche", Voyant_vert => "T_P_VOYANT_VERT", Marche_systeme => "Marche_systeme", Voyant_rouge => "T_P_VOYANT_ROUGE")
   END_RUNG
   RUNG wire#powerrail
      I_Contact( "T_Mode_Manu_VUP" )
   END_RUNG wire#w1
   // the same network as SCL:
   IF NOT "Mode_Manu_Auto" OR NOT "T_Mode_Manu_VUP" THEN
       "Marche_Arret_DB"(Bouton_Rouge := "T_P_Arret",   // "Marche_Arret"
                         Bouton_Vert := "T_P_Marche",
                         Voyant_vert => "T_P_VOYANT_VERT",
                         Marche_systeme => "Marche_systeme",
                         Voyant_rouge => "T_P_VOYANT_ROUGE");
   END_IF;
END_REGION

REGION Network 5: Conduite
   RUNG wire#powerrail
      I_Contact( "Mode_Manu_Auto" )
      wire#w1
      "Conduite_DB"(Marche := "Marche_systeme", Fin_bras := "T_fin_bras_poste_1", Fin_ascenseur := "T_fin_ascenseur", Fin_test_couleur := "T_fin_test_couleur", Fin_test_epaisseur := "T_Fin_test_epaisseur", Fonctionnement_init := "T_fonctionnement_init", présence_pice_mag := "T_Piece_Mag", DEBUT_BRAS => "T_debut_bras", DEBUT_ASCENSEUR => "T_debut_asc", DEBUT_EPAISSEUR => "T_debut_test_epaisseur", DEBUT_TEST_COULEUR => "T_debut_test_couleur", fonctionnement_auto => "T_fonctionnement_auto")
   END_RUNG
   RUNG wire#powerrail
      I_Contact( "T_Mode_Manu_VUP" )
   END_RUNG wire#w1
   // the same network as SCL:
   IF NOT "Mode_Manu_Auto" OR NOT "T_Mode_Manu_VUP" THEN
       "Conduite_DB"(Marche := "Marche_systeme",   // "Conduite"
                     Fin_bras := "T_fin_bras_poste_1",
                     Fin_ascenseur := "T_fin_ascenseur",
                     Fin_test_couleur := "T_fin_test_couleur",
                     Fin_test_epaisseur := "T_Fin_test_epaisseur",
                     Fonctionnement_init := "T_fonctionnement_init",
                     présence_pice_mag := "T_Piece_Mag",
                     DEBUT_BRAS => "T_debut_bras",
                     DEBUT_ASCENSEUR => "T_debut_asc",
                     DEBUT_EPAISSEUR => "T_debut_test_epaisseur",
                     DEBUT_TEST_COULEUR => "T_debut_test_couleur",
                     fonctionnement_auto => "T_fonctionnement_auto");
   END_IF;
END_REGION

REGION Network 6: Bras Poste 1
   RUNG wire#powerrail
      I_Contact( "Mode_Manu_Auto" )
      wire#w1
      "Bras_poste_1_DB"(bras_asc := "T_Bras_Asc", presence_piece := "T_Piece_Mag", marche := "T_debut_bras", bras_mag := "T_Bras_Mag", vide_bon := "T_Vide_Bon", FIN_BRAS_POSTE_1 => "T_fin_bras_poste_1")
   END_RUNG
   RUNG wire#powerrail
      I_Contact( "T_Mode_Manu_VUP" )
   END_RUNG wire#w1
   // the same network as SCL:
   IF NOT "Mode_Manu_Auto" OR NOT "T_Mode_Manu_VUP" THEN
       "Bras_poste_1_DB"(bras_asc := "T_Bras_Asc",   // "Bras_poste_1"
                         presence_piece := "T_Piece_Mag",
                         marche := "T_debut_bras",
                         bras_mag := "T_Bras_Mag",
                         vide_bon := "T_Vide_Bon",
                         FIN_BRAS_POSTE_1 => "T_fin_bras_poste_1");
   END_IF;
END_REGION

REGION Network 7: Ascenceur poste 1
   RUNG wire#powerrail
      I_Contact( "Mode_Manu_Auto" )
      wire#w1
      "Ascenseur_poste_1_DB"(asc_bas := "T_Asc_Bas", presence_piece_asc := "T_Piece_Asc", asc_haut := "T_Asc_Haut", Fin_test_epaisseur := "T_Fin_test_epaisseur", marche := "T_debut_asc", MONTER_ASC => "T_MONT_ASC", DESCENDRE_ASC => "T_DESC_ASC", FIN_ASCENSEUR => "T_fin_ascenseur")
   END_RUNG
   RUNG wire#powerrail
      I_Contact( "T_Mode_Manu_VUP" )
   END_RUNG wire#w1
   // the same network as SCL:
   IF NOT "Mode_Manu_Auto" OR NOT "T_Mode_Manu_VUP" THEN
       "Ascenseur_poste_1_DB"(asc_bas := "T_Asc_Bas",   // "Ascenseur_poste_1"
                              presence_piece_asc := "T_Piece_Asc",
                              asc_haut := "T_Asc_Haut",
                              Fin_test_epaisseur := "T_Fin_test_epaisseur",
                              marche := "T_debut_asc",
                              MONTER_ASC => "T_MONT_ASC",
                              DESCENDRE_ASC => "T_DESC_ASC",
                              FIN_ASCENSEUR => "T_fin_ascenseur");
   END_IF;
END_REGION

REGION Network 8: Test Epaisseur
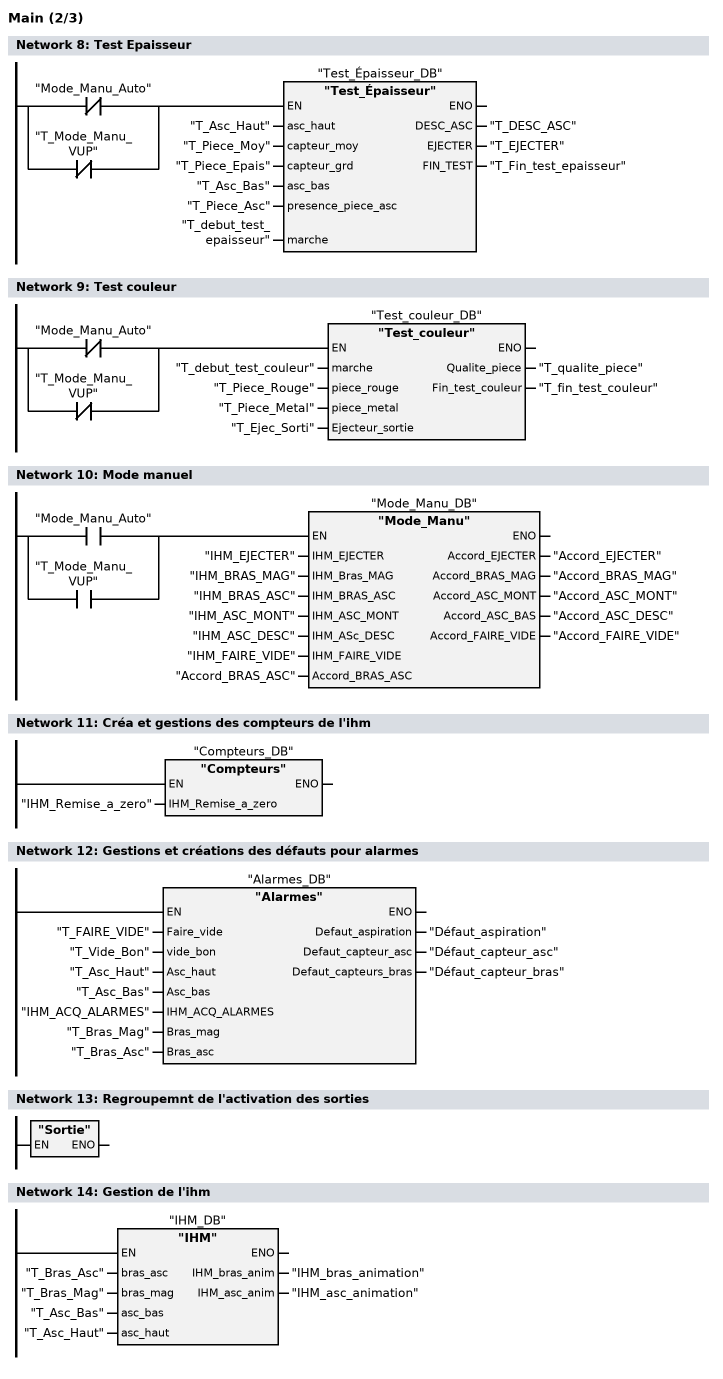
   RUNG wire#powerrail
      I_Contact( "Mode_Manu_Auto" )
      wire#w1
      "Test_Épaisseur_DB"(asc_haut := "T_Asc_Haut", capteur_moy := "T_Piece_Moy", capteur_grd := "T_Piece_Epais", asc_bas := "T_Asc_Bas", presence_piece_asc := "T_Piece_Asc", marche := "T_debut_test_epaisseur", DESC_ASC => "T_DESC_ASC", EJECTER => "T_EJECTER", FIN_TEST => "T_Fin_test_epaisseur")
   END_RUNG
   RUNG wire#powerrail
      I_Contact( "T_Mode_Manu_VUP" )
   END_RUNG wire#w1
   // the same network as SCL:
   IF NOT "Mode_Manu_Auto" OR NOT "T_Mode_Manu_VUP" THEN
       "Test_Épaisseur_DB"(asc_haut := "T_Asc_Haut",   // "Test_Épaisseur"
                           capteur_moy := "T_Piece_Moy",
                           capteur_grd := "T_Piece_Epais",
                           asc_bas := "T_Asc_Bas",
                           presence_piece_asc := "T_Piece_Asc",
                           marche := "T_debut_test_epaisseur",
                           DESC_ASC => "T_DESC_ASC",
                           EJECTER => "T_EJECTER",
                           FIN_TEST => "T_Fin_test_epaisseur");
   END_IF;
END_REGION

REGION Network 9: Test couleur
   RUNG wire#powerrail
      I_Contact( "Mode_Manu_Auto" )
      wire#w1
      "Test_couleur_DB"(marche := "T_debut_test_couleur", piece_rouge := "T_Piece_Rouge", piece_metal := "T_Piece_Metal", Ejecteur_sortie := "T_Ejec_Sorti", Qualite_piece => "T_qualite_piece", Fin_test_couleur => "T_fin_test_couleur")
   END_RUNG
   RUNG wire#powerrail
      I_Contact( "T_Mode_Manu_VUP" )
   END_RUNG wire#w1
   // the same network as SCL:
   IF NOT "Mode_Manu_Auto" OR NOT "T_Mode_Manu_VUP" THEN
       "Test_couleur_DB"(marche := "T_debut_test_couleur",   // "Test_couleur"
                         piece_rouge := "T_Piece_Rouge",
                         piece_metal := "T_Piece_Metal",
                         Ejecteur_sortie := "T_Ejec_Sorti",
                         Qualite_piece => "T_qualite_piece",
                         Fin_test_couleur => "T_fin_test_couleur");
   END_IF;
END_REGION

REGION Network 10: Mode manuel
   RUNG wire#powerrail
      Contact( "Mode_Manu_Auto" )
      wire#w1
      "Mode_Manu_DB"(IHM_EJECTER := "IHM_EJECTER", IHM_Bras_MAG := "IHM_BRAS_MAG", IHM_BRAS_ASC := "IHM_BRAS_ASC", IHM_ASC_MONT := "IHM_ASC_MONT", IHM_ASc_DESC := "IHM_ASC_DESC", IHM_FAIRE_VIDE := "IHM_FAIRE_VIDE", Accord_BRAS_ASC := "Accord_BRAS_ASC", Accord_EJECTER => "Accord_EJECTER", Accord_BRAS_MAG => "Accord_BRAS_MAG", Accord_ASC_MONT => "Accord_ASC_MONT", Accord_ASC_BAS => "Accord_ASC_DESC", Accord_FAIRE_VIDE => "Accord_FAIRE_VIDE")
   END_RUNG
   RUNG wire#powerrail
      Contact( "T_Mode_Manu_VUP" )
   END_RUNG wire#w1
   // the same network as SCL:
   IF "Mode_Manu_Auto" OR "T_Mode_Manu_VUP" THEN
       "Mode_Manu_DB"(IHM_EJECTER := "IHM_EJECTER",   // "Mode_Manu"
                      IHM_Bras_MAG := "IHM_BRAS_MAG",
                      IHM_BRAS_ASC := "IHM_BRAS_ASC",
                      IHM_ASC_MONT := "IHM_ASC_MONT",
                      IHM_ASc_DESC := "IHM_ASC_DESC",
                      IHM_FAIRE_VIDE := "IHM_FAIRE_VIDE",
                      Accord_BRAS_ASC := "Accord_BRAS_ASC",
                      Accord_EJECTER => "Accord_EJECTER",
                      Accord_BRAS_MAG => "Accord_BRAS_MAG",
                      Accord_ASC_MONT => "Accord_ASC_MONT",
                      Accord_ASC_BAS => "Accord_ASC_DESC",
                      Accord_FAIRE_VIDE => "Accord_FAIRE_VIDE");
   END_IF;
END_REGION

REGION Network 11: Créa et gestions des compteurs de l'ihm
   RUNG wire#powerrail
      "Compteurs_DB"(IHM_Remise_a_zero := "IHM_Remise_a_zero")
   END_RUNG
   // the same network as SCL:
   "Compteurs_DB"(IHM_Remise_a_zero := "IHM_Remise_a_zero");   // "Compteurs"
END_REGION

REGION Network 12: Gestions et créations des défauts pour alarmes
   RUNG wire#powerrail
      "Alarmes_DB"(Faire_vide := "T_FAIRE_VIDE", vide_bon := "T_Vide_Bon", Asc_haut := "T_Asc_Haut", Asc_bas := "T_Asc_Bas", IHM_ACQ_ALARMES := "IHM_ACQ_ALARMES", Bras_mag := "T_Bras_Mag", Bras_asc := "T_Bras_Asc", Defaut_aspiration => "Défaut_aspiration", Defaut_capteur_asc => "Défaut_capteur_asc", Defaut_capteurs_bras => "Défaut_capteur_bras")
   END_RUNG
   // the same network as SCL:
   "Alarmes_DB"(Faire_vide := "T_FAIRE_VIDE",   // "Alarmes"
                vide_bon := "T_Vide_Bon",
                Asc_haut := "T_Asc_Haut",
                Asc_bas := "T_Asc_Bas",
                IHM_ACQ_ALARMES := "IHM_ACQ_ALARMES",
                Bras_mag := "T_Bras_Mag",
                Bras_asc := "T_Bras_Asc",
                Defaut_aspiration => "Défaut_aspiration",
                Defaut_capteur_asc => "Défaut_capteur_asc",
                Defaut_capteurs_bras => "Défaut_capteur_bras");
END_REGION

REGION Network 13: Regroupemnt de l'activation des sorties
   RUNG wire#powerrail
      "Sortie"()
   END_RUNG
   // the same network as SCL:
   "Sortie"();
END_REGION

REGION Network 14: Gestion de l'ihm
   RUNG wire#powerrail
      "IHM_DB"(bras_asc := "T_Bras_Asc", bras_mag := "T_Bras_Mag", asc_bas := "T_Asc_Bas", asc_haut := "T_Asc_Haut", IHM_bras_anim => "IHM_bras_animation", IHM_asc_anim => "IHM_asc_animation")
   END_RUNG
   // the same network as SCL:
   "IHM_DB"(bras_asc := "T_Bras_Asc",   // "IHM"
            bras_mag := "T_Bras_Mag",
            asc_bas := "T_Asc_Bas",
            asc_haut := "T_Asc_Haut",
            IHM_bras_anim => "IHM_bras_animation",
            IHM_asc_anim => "IHM_asc_animation");
END_REGION

REGION Network 15: ODDO
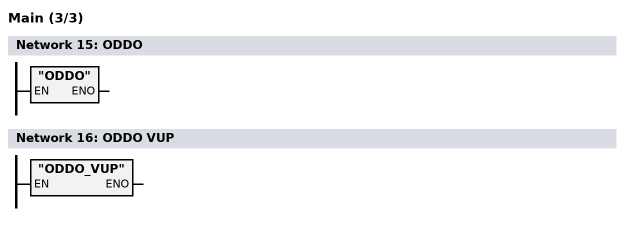
   RUNG wire#powerrail
      "ODDO"()
   END_RUNG
   // the same network as SCL:
   "ODDO"();
END_REGION

REGION Network 16: ODDO VUP
   RUNG wire#powerrail
      "ODDO_VUP"()
   END_RUNG
   // the same network as SCL:
   "ODDO_VUP"();
END_REGION
END_ORGANIZATION_BLOCK

ORGANIZATION_BLOCK "Startup"   // OB100, SCL, Startup
TITLE = "Complete Restart"
{ S7_Optimized_Access := 'TRUE' }
VERSION : 0.1
   VAR_INPUT
      LostRetentive : Bool;   // True if retentive data are lost
      LostRTC : Bool;   // True if date and time are lost
   END_VAR
BEGIN
   //Init des étapes dans grafcets
   "Marche_Arret_DB".Etape_Marche_Arret := 10;
   "Bras_poste_1_DB".Etape_Bras_Poste_1 := 400;
   "Ascenseur_poste_1_DB".Etape_Ascenseur := 500;
   "Test_Épaisseur_DB".Etape_Test_epaisseur := 100;
   "Conduite_DB".Etape_conduite := 1000;
   "Test_couleur_DB".Etape_test_couleur := 700;
   "Initialisation_DB".Etape_init := 2000;

   //Reset des commandes du mode manuel par sécurité
   "Mode_Manu_DB".Accord_ASC_BAS := FALSE;
   "Mode_Manu_DB".Accord_ASC_MONT := FALSE;
   "Mode_Manu_DB".Accord_BRAS_ASC := FALSE;
   "Mode_Manu_DB".Accord_BRAS_MAG := FALSE;
   "Mode_Manu_DB".Accord_EJECTER := FALSE;
   "Mode_Manu_DB".Accord_FAIRE_VIDE := FALSE;

   "Simu_VUP" := FALSE;
END_ORGANIZATION_BLOCK

ORGANIZATION_BLOCK "ProDiagOB"   // OB250, ProDiag_OB, ProgramCycle
TITLE = "Main Program Sweep (Cycle)"
{ S7_Optimized_Access := 'TRUE' }
VERSION : 0.1
   VAR_INPUT
      Initial_Call : Bool;   // Initial call of this OB
      Remanence : Bool;   // =True, if remanent data are available
   END_VAR
BEGIN

REGION Network 1
   CALL "Default_SupervisionFB", "Default_SupervisionDB";
END_REGION
END_ORGANIZATION_BLOCK

// folder: I/O

FUNCTION "IDDI" : Void   // FC1, SCL
{ S7_Optimized_Access := 'TRUE' }
VERSION : 0.1
BEGIN
   IF NOT "Simu_VUP" THEN
       "T_Bras_Asc" := "I_Bras_Asc";
       "T_Bras_Mag" := "I_Bras_Mag";
       "T_Piece_Mag" := "I_Piece_Mag";
       "T_Vide_Bon" := "I_Vide_Bon";
       "T_Piece_Rouge" := "I_Piece_Rouge";
       "T_Piece_Asc" := "I_Piece_Asc";
       "T_Piece_Metal" := "I_Piece_Metal";
       "T_Ejec_Entre" := "I_Ejec_Entre";
       "T_Ejec_Sorti" := "I_Ejec_Sorti";
       "T_Asc_Bas" := "I_Asc_Bas";
       "T_Asc_Haut" := "I_Asc_Haut";
       "T_Piece_Moy" := "I_Piece_Moy";
       "T_Piece_Epais" := "I_Piece_Epais";
       "T_P_Commutateur" := "I_P_Commutateur";
       "T_P_Arret" := "I_P_Arret";
       "T_P_Marche" := "I_P_Marche";
   END_IF;
END_FUNCTION

FUNCTION "ODDO" : Void   // FC2, SCL
{ S7_Optimized_Access := 'TRUE' }
VERSION : 0.1
BEGIN
   IF NOT "Simu_VUP" THEN
       "Q_FAIRE_VIDE" := "T_FAIRE_VIDE";
       "Q_BR_ASC" := "T_BR_ASC";
       "Q_BR_MAG" := "T_BR_MAG";
       "Q_EJECTER" := "T_EJECTER";
       "Q_MONT_ASC" := "T_MONT_ASC";
       "Q_DESC_ASC" := "T_DESC_ASC";

   END_IF;

   "Q_P_VOYANT_ROUGE" := "T_P_VOYANT_ROUGE";
   "Q_P_VOYANT_VERT" := "T_P_VOYANT_VERT";
END_FUNCTION

FUNCTION "ODDO_VUP" : Void   // FC3, SCL
{ S7_Optimized_Access := 'TRUE' }
VERSION : 0.1
BEGIN
   IF "Simu_VUP" = TRUE THEN //20.X
       "Q_VUP_BR_ASC" := "T_BR_ASC";
       "Q_VUP_BR_MAG" := "T_BR_MAG";
       "Q_VUP_FAIRE_VIDE" := "T_FAIRE_VIDE";
       "Q_VUP_EJECTER" := "T_EJECTER";
       "Q_VUP_MONT_ASC" := "T_MONT_ASC";
       "Q_VUP_DESC_ASC" := "T_DESC_ASC";
   END_IF;
END_FUNCTION

FUNCTION "IDDI_VUP" : Void   // FC4, SCL
{ S7_Optimized_Access := 'TRUE' }
VERSION : 0.1
BEGIN
   IF "Simu_VUP" = TRUE THEN //adresse var I_VUP -> 25.x
       "T_Bras_Asc" := "I_VUP_Bras_Asc";
       "T_Bras_Mag" := "I_VUP_Bras_Mag";
       "T_Piece_Mag" := "I_VUP_Piece_MAG";
       "T_Vide_Bon" := "I_VUP_Vide_Bon";

       "T_Asc_Bas" := "I_VUP_Asc_Bas";
       "T_Asc_Haut" := "I_VUP_Asc_Haut";
       "T_Piece_Asc" := "I_VUP_Piece_Asc";

       "T_Piece_Moy" := "I_VUP_Piece_Moy";
       "T_Piece_Epais" := "I_VUP_Piece_Epais";

       "T_P_Arret" := "I_VUP_Arret";
       "T_P_Marche" := "I_VUP_Marche";
       "T_Mode_Manu_VUP" := "I_Mode_Manu_VUP";
   END_IF;
END_FUNCTION

// folder: IHM

FUNCTION_BLOCK "IHM"   // FB14, SCL
{ S7_Optimized_Access := 'TRUE' }
VERSION : 0.1
   VAR_INPUT
      bras_asc : Bool;
      bras_mag : Bool;
      asc_bas : Bool;
      asc_haut : Bool;
   END_VAR
   VAR_OUTPUT
      IHM_bras_anim : Bool;
      IHM_asc_anim : Bool;
   END_VAR
BEGIN
   //Gestion des animations des équipements pour l'ihm


   IF NOT #bras_asc AND NOT #bras_mag THEN
       #IHM_bras_anim := TRUE;
   ELSE
       #IHM_bras_anim := FALSE;
   END_IF;

   IF NOT #asc_bas AND NOT #asc_haut THEN
       #IHM_asc_anim := TRUE;
   ELSE
       #IHM_asc_anim := FALSE;
   END_IF;
END_FUNCTION_BLOCK

// folder: Safety

FUNCTION_BLOCK "Main_Safety_RTG1"   // FB1, F_FBD
{ S7_Optimized_Access := 'TRUE' }
   VAR
      ESTOP1_Instance : ESTOP1;
      Arret_Urgence_Instance : "Arret_Urgence";
   END_VAR
BEGIN

REGION Network 1: Sortie Safety
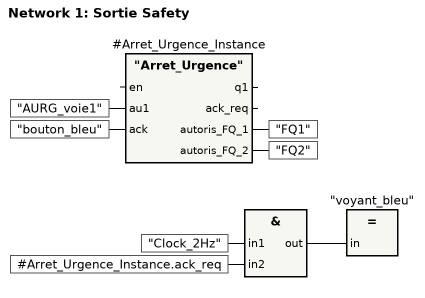
   #Arret_Urgence_Instance(au1 := "AURG_voie1",   // "Arret_Urgence"
                           ack := "bouton_bleu",
                           autoris_FQ_1 => "FQ1",
                           autoris_FQ_2 => "FQ2");
   "voyant_bleu" := "Clock_2Hz" AND #Arret_Urgence_Instance.ack_req;
END_REGION
END_FUNCTION_BLOCK

FUNCTION_BLOCK "Arret_Urgence"   // FB2, F_LAD
{ S7_Optimized_Access := 'TRUE' }
VERSION : 0.1
   VAR_INPUT
      au1 : Bool;
      ack : Bool;
   END_VAR
   VAR_OUTPUT
      q1 : Bool;
      ack_req : Bool;
      autoris_FQ_1 : Bool;
      autoris_FQ_2 : Bool;
   END_VAR
   VAR
      ESTOP1_Instance : ESTOP1;
      sortie_acq_req : ESTOP1;
   END_VAR
   VAR_TEMP   // added for the SCL form of the ladder/FBD networks
      _w1 : Bool;
   END_VAR
BEGIN

REGION Network 1
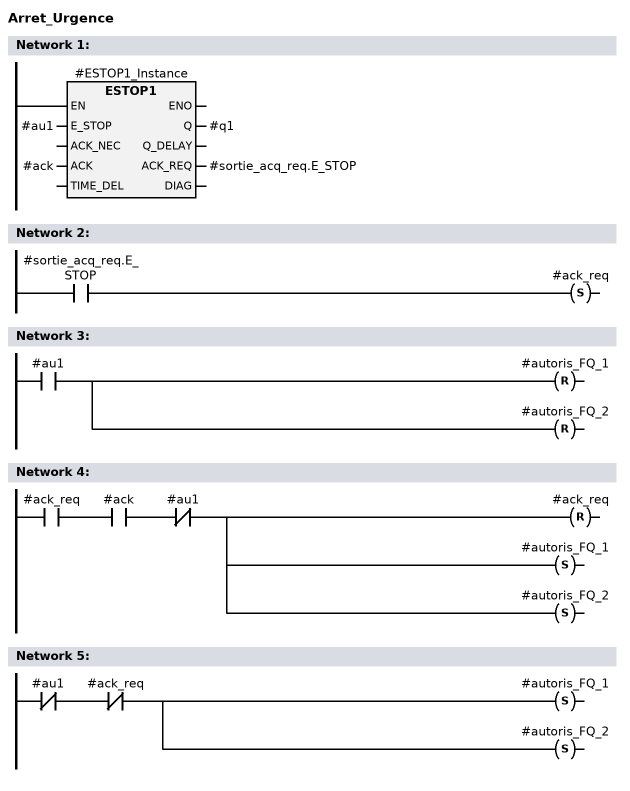
   #ESTOP1_Instance(E_STOP := #au1, ACK := #ack, Q => #q1, ACK_REQ => #sortie_acq_req.E_STOP);   // ESTOP1
END_REGION

REGION Network 2
   RUNG wire#powerrail
      Contact( #sortie_acq_req.E_STOP )
      S_Coil( #ack_req )
   END_RUNG
   // the same network as SCL:
   IF #sortie_acq_req.E_STOP THEN #ack_req := TRUE; END_IF;
END_REGION

REGION Network 3
   RUNG wire#powerrail
      Contact( #au1 )
      wire#w1
      R_Coil( #autoris_FQ_1 )
   END_RUNG
   RUNG wire#w1
      R_Coil( #autoris_FQ_2 )
   END_RUNG
   // the same network as SCL:
   IF #au1 THEN
       #autoris_FQ_1 := FALSE;
       #autoris_FQ_2 := FALSE;
   END_IF;
END_REGION

REGION Network 4
   RUNG wire#powerrail
      Contact( #ack_req )
      Contact( #ack )
      I_Contact( #au1 )
      wire#w1
      R_Coil( #ack_req )
   END_RUNG
   RUNG wire#w1
      S_Coil( #autoris_FQ_1 )
   END_RUNG
   RUNG wire#w1
      S_Coil( #autoris_FQ_2 )
   END_RUNG
   // the same network as SCL:
   #_w1 := #ack_req AND #ack AND NOT #au1;
   IF #_w1 THEN
       #ack_req := FALSE;
       #autoris_FQ_1 := TRUE;
       #autoris_FQ_2 := TRUE;
   END_IF;
END_REGION

REGION Network 5
   RUNG wire#powerrail
      I_Contact( #au1 )
      I_Contact( #ack_req )
      wire#w1
      S_Coil( #autoris_FQ_1 )
   END_RUNG
   RUNG wire#w1
      S_Coil( #autoris_FQ_2 )
   END_RUNG
   // the same network as SCL:
   IF NOT #au1 AND NOT #ack_req THEN
       #autoris_FQ_1 := TRUE;
       #autoris_FQ_2 := TRUE;
   END_IF;
END_REGION
END_FUNCTION_BLOCK

(* ===== HMI "HMI_RT_1" =====
connection "Connexion_1": ETHERNET, ILRT_S7_1500_OMS
connection "HMI_Liaison_1": ETHERNET, ILRT_S7_1500_OMS

HMI tags "Table de variables standard"
   "Numéro_vue" : Int, internal
   "Active_bp_mode_manu" : Bool, internal
   "Active_bp_accueil" : Int, internal
   "Active_bp_Compteur" : Int, internal
   "Active_bp_Alarme" : Int, internal
   "Q_FAIRE_VIDE" : Bool = PLC Q_FAIRE_VIDE AT %Q5.0, T1s
   "Var_Test" : Bool = PLC Var_Test AT %M5.0, T100ms
   "IHM_BRAS_MAG" : Bool = PLC IHM_BRAS_MAG AT %M5.2, T1s
   "IHM_BRAS_ASC" : Bool = PLC IHM_BRAS_ASC AT %M5.1, T1s
   "Mode_Manu_Auto" : Bool = PLC Mode_Manu_Auto AT %M5.5, T1s
   "IHM_ASC_MONT" : Bool = PLC IHM_ASC_MONT AT %M5.3, T1s
   "IHM_ASC_DESC" : Bool = PLC IHM_ASC_DESC AT %M5.4, T1s
   "Simu_VUP" : Bool = PLC Simu_VUP AT %M20.0, T1s
   "IHM_FAIRE_VIDE" : Bool = PLC IHM_FAIRE_VIDE AT %M6.5, T1s
   "IHM_EJECTER" : Bool = PLC IHM_EJECTER AT %M7.0, T1s
   "Compteurs_grande_pièce" : Int = PLC Compteurs_grande_pièce AT %MW8, T1s
   "Compteurs_moyenne_pièce" : Int = PLC Compteurs_moyenne_pièce AT %MW10, T1s
   "Compteurs_petite_pièce" : Int = PLC Compteurs_petite_pièce AT %MW14, T1s
   "IHM_Remise_a_zero" : Bool = PLC IHM_Remise_a_zero AT %M7.1, T1s
   "Compteurs_pièce_noire" : Int = PLC Compteurs_pièce_noire AT %MW16, T1s
   "Compteurs_pièce_rouge" : Int = PLC Compteurs_pièce_rouge AT %MW18, T1s
   "Compteurs_pièce_métal" : Int = PLC Compteurs_pièce_métal AT %MW22, T1s
   "IHM_DEMANDE_INIT" : Bool = PLC IHM_DEMANDE_INIT AT %M7.2, T1s
   "Défaut_aspiration" : Bool = PLC Défaut_aspiration AT %M7.3, T1s
   "Défaut_capteur_asc" : Bool = PLC Défaut_capteur_asc AT %M7.4, T1s
   "Défaut_capteur_bras" : Bool = PLC Défaut_capteur_bras AT %M7.5, T1s
   "IHM_ACQ_ALARMES" : Bool = PLC IHM_ACQ_ALARMES AT %M7.6, T1s
   "T_Bras_Asc" : Bool = PLC T_Bras_Asc AT %M12.0, T1s
   "T_Bras_Mag" : Bool = PLC T_Bras_Mag AT %M12.1, T1s
   "T_Asc_Bas" : Bool = PLC T_Asc_Bas AT %M13.1, T1s
   "T_Asc_Haut" : Bool = PLC T_Asc_Haut AT %M13.2, T1s
   "T_Ejec_Sorti" : Bool = PLC T_Ejec_Sorti AT %M13.0, T1s
   "T_FAIRE_VIDE" : Bool = PLC T_FAIRE_VIDE AT %M4.0, T1s
   "T_Piece_Mag" : Bool = PLC T_Piece_Mag AT %M12.2, T1s
   "T_Piece_Asc" : Bool = PLC T_Piece_Asc AT %M12.5, T1s
   "Compteurs_pièce_total" : Int = PLC Compteurs_pièce_total AT %MW26, T1s
   "T_P_VOYANT_VERT" : Bool = PLC T_P_VOYANT_VERT AT %M5.7, T1s
   "T_P_VOYANT_ROUGE" : Bool = PLC T_P_VOYANT_ROUGE AT %M5.6, T1s
   "IHM_asc_animation" : Bool = PLC IHM_asc_animation AT %M20.6, T1s
   "IHM_bras_animation" : Bool = PLC IHM_bras_animation AT %M7.7, T1s
   "IHM_RESET_INIT" : Bool = PLC IHM_RESET_INIT AT %M20.7, T1s
   "T_fonctionnement_auto" : Bool = PLC T_fonctionnement_auto AT %M4.6, T1s

discrete alarms
   1: 'Défaut du vide, aspiration en cours sans réussite', class Alarm, trigger "Défaut_aspiration" bit 0
   2: 'Défaut des capteurs de position de l'ascenseur', class Alarm, trigger "Défaut_capteur_asc" bit 0
   3: 'Défaut des capteurs de positions du bras', class Alarm, trigger "Défaut_capteur_bras" bit 0

text list "SystemTextList_ConfigErrorAlarmTextLibrary_1": 1 'Erreur de configuration NameService : Suppression implicite. L'instance de sous-élément @6%s@ doit être supprimée explicitement.'; 2 'Erreur de configuration NameService : Suppression implicite. L'instance d'alias/format/unité @6%s@ doit être supprimée explicitement.'

text list "SystemTextList_ConfigErrorAlarmTextLibrary_2": 1 'EvDpManager::cleanupDeletedDatapoint - alert handler config is deleted implicitly for deleted datapoint, @3%s@'; 2 'EvDpManager::cleanupDeletedDatapoint - alert handler config is deleted implicitly but still has overrides, @3%s@'; 3 'EvDpManager::cleanupDeletedDatapoint - default value config is deleted implicitly for deleted datapoint, @3%s@'; 4 'EvDpManager::cleanupDeletedDatapoint - default value config is deleted implicitly but still has overrides, @3%s@'; 5 'EvDpManager::cleanupDeletedDatapoint - initial value config is deleted implicitly for deleted datapoint, @3%s@'; 6 'EvDpManager::cleanupDeletedDatapoint - initial value config is deleted implicitly but still has overrides, @3%s@'; 7 'EvDpManager::cleanupDeletedDatapoint - distribution config is deleted implicitly for deleted datapoint, @3%s@'; 8 'EvDpManager::cleanupDeletedDatapoint - distribution config is deleted implicitly but still has overrides, @3%s@'; 9 'EvDpManager::cleanupDeletedDatapoint - rangeCheck config is deleted implicitly for deleted datapoint, @3%s@'; 10 'EvDpManager::cleanupDeletedDatapoint - rangeCheck config is deleted implicitly but still has overrides, @3%s@'

text list "SystemTextList_ConfigErrorAlarmTextLibrary_3": 1 'Le type de point de données configuré a été supprimé, mais un type configuré est encore défini pour le type de noeud : @3%s@.'; 2 'Le type de noeud de point de données configuré a été supprimé dans le type de point de données, mais un type configuré est encore défini pour l'élément : @3%s@.'

text list "SystemTextList_ConfigErrorAlarmTextLibrary_4": 2 'Cycles : @6%s@ n'existe pas.'; 3 'Alarmes : @6%s@ existe déjà.'; 4 'Variables : L'adresse @6%s@ a été rejetée.'; 1 'Connexions : @6%s@ n'existe pas.'; 5 'Variables : Le mode d'acquisition @6%s@ n'est pas pris en charge.'; 6 'Cycles : @6%s@ a été supprimé, mais des variables associées existent.'; 7 'Connexions : @6%s@ a été supprimé, mais des variables associées existent.'; 8 'Variables : La variable @6%s@ a été rejetée.'; 9 'Variables : La variable @6%s@ a une valeur invalide.'; 10 'Les adresses multiplex ne sont pas autorisées pour la configuration de tableaux de bloc (nom DP : @3%s@)'; 11 'La configuration de tableau de bloc est erronée (nom DP : @3%s@)'; 12 'La configuration de tableau de bloc n'est pas prise en charge par le système redondant (nom DP : @3%s@)'; 13 'Les variables Tableau de bloc ne sont pas prises en charge par l'adaptateur de protocole (nom DP : @3%s@)'; 14 'L'adresse de périphérie de la variable Handshake Tableau de bloc n'existe pas (nom DP : @3%s@)'; 15 'Le nombre de configurations de tableau de bloc dépasse le nombre maximum (<@6%s@)'; 16 'Le nombre d'éléments des configurations de tableau de bloc dépasse le nombre maximum (nom DP : @3%s@, taille : @6%s@)'; 17 'Variable Handshake qui est référencée par plusieurs configurations de tableau de bloc (nom DP : @3%s@)'; 0 'Connexions : Impossible d'établir la connexion à @6%s@'; 65638 'Connexions : Impossible d'établir la connexion à @6%s@'; 65639 'Connexions : @6%s@ coupée'; 65640 'Connexions : Connexion à l'appareil IHM @6%s@ coupée'; 65641 'Connexions : Connexion à l'API @6%s@ coupée'; 65541 'Connexions : Dépassement de temps lors de l'établissement de la connexion à @6%s@'; 65542 'Connexions : perturbé - @5%s@'; 65543 'Connexions : Connexion à l'appareil IHM coupée. La connexion @5%s@ a été modifiée.'; 65544 'Connexions : Connexion à l'appareil IHM coupée. La propriété du pilote a été modifiée pour la connexion @5%s@.'

text list "SystemTextList_ConfigErrorAlarmTextLibrary_5": 1 'Connexions : Le cycle de la surveillance de signe de vie doit être inférieur au temps de réponse.'; 2 'Connexions : Des services cycliques sont configurés, mais ne sont pas pris en charge par l'appareil cible.'; 3 'Connexions : Une lecture sur modification est configurée, mais n'est pas prise en charge par l'appareil cible.'; 4 'Variables : L'adresse @6%s@ n'existe pas dans l'API.'; 5 'Variables : Impossible de déterminer le type de conversion par défaut pour l'adresse @6%s@.'; 6 'Variables : Type de conversion invalide'; 7 'Cycles : Type de conversion invalide. La conversion n'est pas prise en charge sur le cycle HmiCycle.'; 4096 'Connexions : La version de l'adresse @6%s@ n'est pas prise en charge.'; 4097 'Connexions : L'adresse Profibus n'est pas prise en charge.'; 4098 'Connexions : L'adresse Softbus n'est pas prise en charge.'; 4099 'Connexions : Le type d'adresse @6%s@ n'est pas pris en charge.'; 4100 'Connexions : Connexion nommée invalide @6%s@. Le point d'accès n'est pas pris en compte.'; 4101 'Connexions : Le routage n'est pas pris en charge. @6%s@ ne sera pas utilisé.'; 4102 'Connexions : Le routage n'est pas pris en charge. @6%s@ ne sera pas utilisé.'; 4103 'Connexions : Adresse IP invalide @6%s@'; 4104 'Connexions : Connexion nommée invalide @6%s@. Format valide : >VMD</>connexion<'; 4105 'Connexions : Connexion nommée invalide @6%s@. Le nom de connexion VMD est trop long. 24 caractères sont autorisés au plus.'; 4106 'Connexions : Connexion nommée invalide @6%s@. Le nom de connexion est trop long. 32 caractères sont autorisés au plus.'; 4107 'Connexions : Le numéro de châssis @6%s@ se situe hors de la plage autorisée (0..7).'; 4108 'Connexions : Connexion nommée invalide @6%s@. Le châssis n'est pas pris en compte.'; 4109 'Connexions : Le numéro d'emplacement @6%s@ se situe hors de la plage autorisée (0..31)'; 4110 'Connexions : Connexion nommée invalide @6%s@. L'emplacement n'est pas pris en compte.'; 4111 'Impossible d'établir la connexion. Le nombre maximum de connexions disponibles (@6%s@) est dépassé.'; 4112 'Connexion coupée. Aucun signe de vie pendant les @4%s@ dernières ms.'; 4113 'Impossible d'établir la connexion - @4%s@'; 4114 'Impossible d'établir la connexion. L'adresse @6%s@ n'est pas utilisable.'; 4115 'Impossible d'établir la connexion. Adresse invalide @6%s@'; 4116 'Impossible d'établir la connexion - @4%s@'

text list "SystemTextList_ConfigErrorAlarmTextLibrary_6": 1 'Impossible d'établir la connexion. Le certificat d'instance d'application n'est pas configuré.'; 2 'Impossible d'établir la connexion. Le serveur a rejeté le certificat client. Code d'état OPC UA @4%s@'; 3 'Impossible d'établir la connexion. Problème interne dans le magasin de certificats. Code d'état OPC UA @4%s@'; 4 'Impossible d'établir la connexion. Le certificat d'instance d'application n'a pas pu être chargé. Code d'état OPC UA @4%s@'; 5 'Impossible d'établir la connexion. Le serveur n'a pas fourni de certificat. @4%s@'; 6 'Impossible d'établir la connexion. La validation du certificat du serveur a échoué. Code d'état OPC UA @4%s@'; 7 'La connexion a été fermée. Erreur lors de la synchronisation des alarmes. Code d'état OPC UA @4%s@'; 8 'La connexion a été fermée. L'abonnement aux alarmes/événements a échoué. Le nombre d'opérations sur le serveur a été dépassé.'; 9 'La connexion a été fermée. L'abonnement aux alarmes/événements a échoué. Le nombre d'abonnements aux alarmes/événements sur le serveur a été dépassé.'; 10 'Impossible d'établir la connexion. Le serveur signale un problème de licence. Code d'état OPC UA @4%s@'; 11 'Impossible d'établir la connexion. Le nombre maximum de sessions sur le serveur a été dépassé.'; 12 'Impossible d'établir la connexion. La configuration de sécurité est incohérente. @4%s@'; 13 'Impossible d'établir la connexion. L'adresse @4%s@ n'est pas utilisable.'; 14 'Impossible d'établir la connexion. Code d'état OPC UA @4%s@'; 15 'Connexion coupée. Le serveur OPC UA a été arrêté.'; 16 'Connexion coupée. Aucun signe de vie pendant les @4%s@ dernières ms.'; 17 'La connexion a été fermée. Maintenance du serveur OPC UA'; 18 'Impossible d'établir la connexion. Configuration invalide du mode d'authentification. @4%s@'; 19 'Impossible d'établir la connexion. L'utilisateur n'a pas pu être authentifié. Code d'état OPC UA @4%s@'; 20 'Impossible d'établir la connexion. Le serveur n'autorise pas les connexions anonymes. Code d'état OPC UA @4%s@'; 21 'Impossible d'établir la connexion. Problème de certificat : erreur lors de l'écriture des données de sécurité dans @4%s@'; 22 'Impossible d'établir la connexion. Problème de certificat : impossible de supprimer un fichier inattendu dans le répertoire @4%s@'; 23 'Impossible d'établir la connexion. L'utilisateur n'a pas pu être authentifié. Aucun utilisateur ou mot de passe n'est configuré.'; 24 'Impossible d'établir la connexion. Longueur inattendue du certificat du serveur. @4%s@'; 25 'Impossible d'établir la connexion. @4%s@ sans contenu'; 26 'Impossible d'établir la connexion. @4%s@ a un format inattendu.'; 27 'Impossible d'établir la connexion. Les points finaux du serveur ne peuvent pas être lus. Code d'état OPC UA @4%s@'; 28 'Impossible d'établir la connexion. Les points finaux du serveur sont introuvables. @4%s@'; 29 'Impossible d'établir la connexion. Le certificat d'instance d'application est introuvable.'; 30 'Impossible d'établir la connexion. Format inattendu du certificat @4%s@'; 31 'Impossible d'établir la connexion. Format inattendu de la liste de révocation des certificats @4%s@'; 32 'Impossible d'établir la connexion. L'utilisateur n'a pas pu être authentifié. Un détail de cryptage est invalide. @4%s@'; 34 'Impossible d'établir la connexion. - Le mode de redondance non transparent configuré @4%s@ n'est pas pris en charge.'; 101 'Variables : L'adresse @6%s@ n'existe pas sur le serveur.'; 103 'Variables : Impossible d'accéder à l'adresse @6%s@'; 104 'Variables : Le mode d'acquisition n'est pas pris en charge pour l'adresse @6%s@.'; 201 'Alarmes : L'adresse @6%s@ n'existe pas sur le serveur.'; 202 'Alarmes : Impossible d'utiliser l'adresse @6%s@. Le filtre de zone indiqué n'est pas un Event Notifier OPC UA.'; 203 'Alarmes : Impossible d'utiliser l'adresse @6%s@. Le filtre de zone indiqué n'existe pas sur le serveur.'; 204 'Alarmes : Impossible d'utiliser l'adresse @6%s@, car il ne s'agit pas d'un type d'événement OPC UA.'; 205 'Alarmes : Impossible d'utiliser l'adresse @6%s@, car le type de condition OPC UA n'est pas pris en charge.'; 206 'Alarmes : Impossible d'utiliser l'adresse @6%s@, car le type d'événement n'existe pas sur le serveur.'; 207 'Alarmes : Impossible d'utiliser le mode d'acquisition pour l'adresse @6%s@'; 301 'Impossible d'utiliser l'adresse @6%s@, car le numéro de version manque.'; 302 'Impossible d'utiliser l'adresse @6%s@, car le numéro de version est invalide.'; 303 'Impossible d'utiliser l'adresse @6%s@, car le nombre de séparateurs '$' est invalide.'; 304 'Impossible d'utiliser l'adresse @6%s@, car le type d'adresse est invalide.'; 305 'Version non prise en charge @6%s@ de l'adresse'; 401 'Réponse inattendue du serveur OPC UA : @6%s@'

text list "SystemTextList_ConfigErrorAlarmTextLibrary_7": 1 'Alarmes : Chaîne de condition invalide pour l'affichage d'alarme @6%s@'; 2 'Alarmes : Variable et bit d'état invalides pour l'affichage d'alarme @6%s@'; 3 'Alarmes : Variable et bit de commande invalides pour l'affichage d'alarme @6%s@'

text list "SystemTextList_ConfigErrorAlarmTextLibrary_8": 1 'Archives : Suppression implicite. L'instance de variable d'archive @6%s@ doit être supprimée, mais il existe des éléments prioritaires.'

text list "SystemTextList_ConfigErrorAlarmTextLibrary_9": 2 'Un redémarrage du runtime est nécessaire.'; 3 'Il faut éjecter puis ré-insérer le support de stockage correct.'

text list "SystemTextList_ConfigErrorAlarmTextLibrary_10": 1 'Cache CDS : Impossible de créer le répertoire cache ou d'y accéder : @6%s@'; 2 'Cache LOC : Impossible de créer le répertoire cache ou d'y accéder : @6%s@'

text list "SystemTextList_RuntimeCollaborationFailureReason_1": 0 'Erreur inconnue (@3%s@)'; 1 'Le système ne fonctionne pas ou il y a un problème de réseau'; 2 'Runtime n'est pas démarré sur le système cible.'; 3 'L'ID système ne correspond pas à l'ID système attendue @3%s@'; 4 'Le nom de Collaboration ne correspond pas au nom de Collaboration attendu "@3%s@"'; 5 'Certificat erroné ou inconnu'; 6 'Certificat révoqué'; 7 'La différence de temps est trop grande.'; 8 'No common supported message version'; 9 'L'ID système (@3%s@) existe déjà'; 10 'Le nom système (@3%s@) existe déjà'; 11 'ID/Nom existe déjà dans la configuration locale pour Runtime Collaboration'; 12 'L'ID système est en conflit avec une connexion configurée localement (@3%s@)'; 13 'Le nom système est en conflit avec une connexion configurée localement (@3%s@)'

text list "SystemTextList_RedundancyRecoveryFailureReason_1": 0 'Demande de restauration des données temporairement rejetée, jusqu'à ce qu'une réponse soit apportée à la demande de restauration propre.'; 1 'Demande de restauration des données rejetée. Sauvegarde en ligne en cours.'; 2 'Demande de restauration des données rejetée. La connexion au gestionnaire d'événements n'est pas établie.'; 3 'Demande de restauration des données temporairement rejetée jusqu'à l'achèvement de l'activation des modifications.'; 4 'Demande de restauration des données temporairement rejetée tant que les alarmes et les variables persistent.'; 5 'Demande de restauration des données refusée. Le fichier obligatoire config.level.es est manquant sur l'ordinateur.'; 6 'La demande de restauration des données a été annulée par le gestionnaire d'événements.'; 7 'Échec de la synchronisation des données entre les appareils.'; 8 'Différents projets sont démarrés sur les ordinateurs.'

text list "SystemTextList_S7PlusAlarmTextListCollection_1": 4096 'Connexions : Connexion à l'API coupée - @4%s@'; 4097 'Connexions : Connexion à l'appareil IHM coupée - @4%s@'; 4098 'Nombre maximal de liaisons dépassé - @4%s@'; 4099 'Ressources disponibles insuffisantes sur l'API - @4%s@'; 4100 'Échec de légitimation, mot de passe erroné ou manquant - @4%s@'; 4101 'Échec de la demande de liaison pour l'ouverture de la liaison - @4%s@'; 4102 'Connexions : Échec de l'ouverture de la liaison à l'API - @4%s@'; 4103 'Impossible d'envoyer la demande de liaison pour l'ouverture de la liaison'; 4104 'Erreur de certificat générale pour API - @4%s@'; 4105 'Le certificat API a expiré pour - @4%s@'; 4106 'Le certificat API est verrouillé pour - @4%s@'; 4107 'Le certificat API n'est pas de confiance. L'attribution manuelle de la confiance est possible pour - @4%s@'; 4108 'Le certificat API n'est pas de confiance. L'attribution manuelle de la confiance n'est pas possible pour - @4%s@'

text list "SystemTextList_AllenBradleyEIPAlarmTextListCollection_7": 4096 'Liaison perdue côté API - @5%s@'; 4097 'Liaison perdue côté IHM - @5%s@'; 4098 'Nombre maximal de liaisons dépassé - @5%s@'; 4099 'Ressources disponibles insuffisantes sur l'API - @5%s@'; 4100 'Échec de légitimation, mot de passe erroné ou manquant - @5%s@'; 4101 'Échec de la demande de liaison pour l'ouverture de la liaison - @5%s@'; 4102 'Échec de l'ouverture de la liaison - @5%s@'; 4103 'Impossible d'envoyer la demande de liaison pour l'ouverture de la liaison'; 4104 'root certificate expired for - @5%s@'; 4105 'PLC certificate untrusted for - @5%s@'

text list "SystemTextList_AllenBradleyDF1AlarmTextListCollection_9": 4096 'Connexions : Connexion à l'API @5%s@ coupée'; 4097 'Connexions : Connexion à l'appareil IHM @5%s@ coupée'; 4098 'Nombre maximal de liaisons dépassé - @5%s@'; 4099 'Ressources disponibles insuffisantes sur l'API - @5%s@'; 4100 'Échec de légitimation, mot de passe erroné ou manquant - @5%s@'; 4101 'Échec de la demande de liaison pour l'ouverture de la liaison - @5%s@'; 4102 'Connexions : Échec de l'ouverture de la liaison - @5%s@'; 4103 'Impossible d'envoyer la demande de liaison pour l'ouverture de la liaison'; 4104 'Erreur de certificat générale pour API - @5%s@'; 4105 'Le certificat API a expiré pour - @5%s@'; 4106 'Le certificat API est verrouillé pour - @5%s@'; 4107 'Le certificat API n'est pas de confiance. L'attribution manuelle de la confiance est possible pour - @5%s@'; 4108 'Le certificat API n'est pas de confiance. L'attribution manuelle de la confiance n'est pas possible pour - @5%s@'

text list "SystemTextList_OmronEIPAlarmTextListCollection_6": 4096 'Liaison perdue côté API - @5%s@'; 4097 'Liaison perdue côté IHM - @5%s@'; 4098 'Nombre maximal de liaisons dépassé - @5%s@'; 4099 'Ressources disponibles insuffisantes sur l'API - @5%s@'; 4100 'Échec de légitimation, mot de passe erroné ou manquant - @5%s@'; 4101 'Échec de la demande de liaison pour l'ouverture de la liaison - @5%s@'; 4102 'Échec de l'ouverture de la liaison - @5%s@'; 4103 'Impossible d'envoyer la demande de liaison pour l'ouverture de la liaison'; 4104 'root certificate expired for - @5%s@'; 4105 'PLC certificate untrusted for - @5%s@'

text list "SystemTextList_StdModbusTCPAlarmTextListCollection_5": 4096 'Connexions : Connexion à l'API @5%s@ coupée'; 4097 'Connexions : Connexion à l'appareil IHM @5%s@ coupée'; 4098 'Nombre maximal de liaisons dépassé - @5%s@'; 4099 'Ressources disponibles insuffisantes sur l'API - @5%s@'; 4100 'Échec de légitimation, mot de passe erroné ou manquant - @5%s@'; 4101 'Échec de la demande de liaison pour l'ouverture de la liaison - @5%s@'; 4102 'Connexions : Échec de l'ouverture de la liaison - @5%s@'; 4103 'Impossible d'envoyer la demande de liaison pour l'ouverture de la liaison'; 4104 'Erreur de certificat générale pour API - @5%s@'; 4105 'Le certificat API a expiré pour - @5%s@'; 4106 'Le certificat API est verrouillé pour - @5%s@'; 4107 'Le certificat API n'est pas de confiance. L'attribution manuelle de la confiance est possible pour - @5%s@'; 4108 'Le certificat API n'est pas de confiance. L'attribution manuelle de la confiance n'est pas possible pour - @5%s@'

text list "SystemTextList_MitsubishiMCAlarmTextListCollection_4": 4096 'Liaison perdue côté API - @5%s@'; 4097 'Liaison perdue côté IHM - @5%s@'; 4098 'Nombre maximal de liaisons dépassé - @5%s@'; 4099 'Ressources disponibles insuffisantes sur l'API - @5%s@'; 4100 'Échec de légitimation, mot de passe erroné ou manquant - @5%s@'; 4101 'Échec de la demande de liaison pour l'ouverture de la liaison - @5%s@'; 4102 'Échec de l'ouverture de la liaison - @5%s@'; 4103 'Impossible d'envoyer la demande de liaison pour l'ouverture de la liaison'; 4104 'root certificate expired for - @5%s@'; 4105 'PLC certificate untrusted for - @5%s@'

text list "SystemTextList_MitsubishiiQAlarmTextListCollection_3": 4096 'Liaison perdue côté API - @5%s@'; 4097 'Liaison perdue côté IHM - @5%s@'; 4098 'Nombre maximal de liaisons dépassé - @5%s@'; 4099 'Ressources disponibles insuffisantes sur l'API - @5%s@'; 4100 'Échec de légitimation, mot de passe erroné ou manquant - @5%s@'; 4101 'Échec de la demande de liaison pour l'ouverture de la liaison - @5%s@'; 4102 'Échec de l'ouverture de la liaison - @5%s@'; 4103 'Impossible d'envoyer la demande de liaison pour l'ouverture de la liaison'; 4104 'root certificate expired for - @5%s@'; 4105 'PLC certificate untrusted for - @5%s@'

text list "SystemTextList_StdModbusRTUAlarmTextListCollection_8": 4096 'Connexions : Connexion à l'API @5%s@ coupée'; 4097 'Connexions : Connexion à l'appareil IHM @5%s@ coupée'; 4098 'Nombre maximal de liaisons dépassé - @5%s@'; 4099 'Ressources disponibles insuffisantes sur l'API - @5%s@'; 4100 'Échec de légitimation, mot de passe erroné ou manquant - @5%s@'; 4101 'Échec de la demande de liaison pour l'ouverture de la liaison - @5%s@'; 4102 'Connexions : Échec de l'ouverture de la liaison - @5%s@'; 4103 'Impossible d'envoyer la demande de liaison pour l'ouverture de la liaison'; 4104 'Erreur de certificat générale pour API - @5%s@'; 4105 'Le certificat API a expiré pour - @5%s@'; 4106 'Le certificat API est verrouillé pour - @5%s@'; 4107 'Le certificat API n'est pas de confiance. L'attribution manuelle de la confiance est possible pour - @5%s@'; 4108 'Le certificat API n'est pas de confiance. L'attribution manuelle de la confiance n'est pas possible pour - @5%s@'

text list "SystemTextList_LogoAlarmTextListCollection_10": 4096 'Connexions : Connexion à l'API @5%s@ coupée'; 4097 'Connexions : Connexion à l'appareil IHM @5%s@ coupée'; 4098 'Nombre maximal de liaisons dépassé - @5%s@'; 4099 'Ressources disponibles insuffisantes sur l'API - @5%s@'; 4100 'Échec de légitimation, mot de passe erroné ou manquant - @5%s@'; 4101 'Échec de la demande de liaison pour l'ouverture de la liaison - @5%s@'; 4102 'Connexions : Échec de l'ouverture de la liaison - @5%s@'; 4103 'Impossible d'envoyer la demande de liaison pour l'ouverture de la liaison'; 4104 'Erreur de certificat générale pour API - @5%s@'; 4105 'Le certificat API a expiré pour - @5%s@'; 4106 'Le certificat API est verrouillé pour - @5%s@'; 4107 'Le certificat API n'est pas de confiance. L'attribution manuelle de la confiance est possible pour - @5%s@'; 4108 'Le certificat API n'est pas de confiance. L'attribution manuelle de la confiance n'est pas possible pour - @5%s@'

text list "Page_en_cours": 0 'Principale'; 10 'Mode Manu'; 20 'Alarmes'; 30 'Compteurs'
*)

(* ===== HMI "HMI_RT_1" =====

ScreenModuleEditorView "Bloc d'affichage_1" 640x480
   Button "Bouton_1" at 189,135 size 165x65; TextOff 'Text'
*)

(* ===== HMI "HiddenHmiRTDeviceFaceplateTypes" =====

HMI tags "Table de variables standard"
   "TEXT" : Real, internal

HMI tags "b18dabb3-60cf-4a71-8646-bdaaadeb651d"
   "Variable_interface_1" : Real, internal
*)

(* ===== HMI "HiddenHmiRTDeviceFaceplateTypes" =====

HMI tags "Table de variables standard"
   "TEXT" : Real, internal

HMI tags "b18dabb3-60cf-4a71-8646-bdaaadeb651d"
   "Variable_interface_1" : Real, internal
*)

(* ===== HMI "HiddenHmiRTDeviceFaceplateTypes" =====

HMI tags "Table de variables standard"
   "TEXT" : Real, internal

HMI tags "b18dabb3-60cf-4a71-8646-bdaaadeb651d"
   "Variable_interface_1" : Real, internal
*)

(* ===== HMI "HiddenHmiRTDeviceFaceplateTypes" =====

HMI tags "Table de variables standard"
   "TEXT" : Real, internal

HMI tags "b18dabb3-60cf-4a71-8646-bdaaadeb651d"
   "Variable_interface_1" : Real, internal
*)

(* ===== HMI "HiddenHmiRTDeviceFaceplateTypes" =====

HMI tags "Table de variables standard"
   "TEXT" : Real, internal

HMI tags "b18dabb3-60cf-4a71-8646-bdaaadeb651d"
   "Variable_interface_1" : Real, internal
*)

(* ===== HMI "HiddenHmiRTDeviceFaceplateTypes" =====

HMI tags "Table de variables standard"
   "TEXT" : Real, internal

HMI tags "b18dabb3-60cf-4a71-8646-bdaaadeb651d"
   "Variable_interface_1" : Real, internal
*)

(* ===== HMI "HiddenHmiRTDeviceFaceplateTypes" =====

HMI tags "Table de variables standard"
   "TEXT" : Real, internal

HMI tags "b18dabb3-60cf-4a71-8646-bdaaadeb651d"
   "Variable_interface_1" : Real, internal
*)

(* ===== HMI "HiddenHmiRTDeviceFaceplateTypes" =====

HMI tags "Table de variables standard"
   "TEXT" : Real, internal

HMI tags "b18dabb3-60cf-4a71-8646-bdaaadeb651d"
   "Variable_interface_1" : Real, internal
*)

(* ===== HMI "HiddenHmiRTDeviceFaceplateTypes" =====

HMI tags "Table de variables standard"
   "TEXT" : Real, internal

HMI tags "b18dabb3-60cf-4a71-8646-bdaaadeb651d"
   "Variable_interface_1" : Real, internal
*)

(* ===== HMI "HiddenHmiRTDeviceFaceplateTypes" =====

HMI tags "Table de variables standard"
   "TEXT" : Real, internal

HMI tags "b18dabb3-60cf-4a71-8646-bdaaadeb651d"
   "Variable_interface_1" : Real, internal
*)